                                 IF LEN(#mqttTopic) = #LEN_NULL THEN
                                   #statStatus := #ERR_MQTT_COMMAND_UNSUBSCRIBE_TOPIC_INVALID; // Set correct status that identifies error clearly
                                   #statSubfunctionStatus := #ERR_MQTT_COMMAND_UNSUBSCRIBE_TOPIC_INVALID; // Status or return value of called FBs, FCs and system blocks
                                   #statFBErrorState := #statFBState; // Set error state number for diagnostic 
                                   #statErrorUserCleared := TRUE;
                                 ELSE // All ok
                                   //Add two Byte for Paket ID:
                                   #statSendPaketTotalRemLen := #statSendPaketTotalRemLen + #TWO_BYTE_LEN_INFO;
                                   //add unsubscribe  topic len
                                   FOR #tempLoopCounter := #FIRST_CHARACTER TO LEN(#mqttTopic) DO
                                     "LMQTT_ConvertToUtf8"(character     := #mqttTopic[#tempLoopCounter],
                                                           convertedUtf8 => #tempConvertedUtf8,
                                                           bytesUsed     => #tempBytesUsedUtf8,
                                                           error         => #tempErrorConvertUtf8,
                                                           status        => #tempStatusConvertUtf8);
                                     #statUnsubscribeTopicLenUtf8Encoded := #statUnsubscribeTopicLenUtf8Encoded + #tempBytesUsedUtf8;
                                   END_FOR;
                                   //Add len of topic plus len info
                                   #statSendPaketTotalRemLen := #statSendPaketTotalRemLen + #statUnsubscribeTopicLenUtf8Encoded + #TWO_BYTE_LEN_INFO;

                                   //Build Subscribe Telegram
                                   //Fixed Header - Write Paket Type
                                   #statSendBuffer[#statSendBufferPos] := #MQTT_MSG_TYPE_UNSUBSCRIBE;
                                   #statSendBufferPos += 1; // increment

                                   //Write Remaining Paket Len info 
                                   WHILE (#statSendPaketTotalRemLen > #DEFAULT_VALUE_ZERO)
                                   DO//See MQTT Spec for explanation of this calculation
                                     #statEncodedRemPaketLenAsByte := UDINT_TO_BYTE(#statSendPaketTotalRemLen MOD #SEND_LEN_MULTIPLIER_UDINT_128);
                                     #statSendPaketTotalRemLen := #statSendPaketTotalRemLen / #SEND_LEN_MULTIPLIER_UDINT_128;
                                     // if there are more data to encode, set the top bit of this byte
                                     IF #statSendPaketTotalRemLen > #DEFAULT_VALUE_ZERO
                                     THEN
                                       // Do this and continue while loop
                                       #statEncodedRemPaketLenAsByte := #statEncodedRemPaketLenAsByte OR UDINT_TO_BYTE(#SEND_LEN_MULTIPLIER_UDINT_128);
                                       #statSendBuffer[#statSendBufferPos] := #statEncodedRemPaketLenAsByte;
                                       #statSendBufferPos += 1;
                                     ELSE
                                       //do this and leave while loop
                                       #statSendBuffer[#statSendBufferPos] := #statEncodedRemPaketLenAsByte;
                                       #statSendBufferPos += 1;
                                     END_IF;
                                   END_WHILE;

                                   // Set Paket Id
                                   #tempWordForSliceAddress := UINT_TO_WORD(#statPaketId);
                                   #statSendBuffer[#statSendBufferPos] := #tempWordForSliceAddress.%B1; //MSB
                                   #statSendBufferPos += 1;
                                   #statSendBuffer[#statSendBufferPos] := #tempWordForSliceAddress.%B0; //LSB
                                   #statSendBufferPos += 1;

                                   //When all done, set encode to true
                                   #statPaketHeaderEncodeDone := TRUE;
                                 END_IF;
                               END_IF;

                               //Header Encoded - 
                               IF #statPaketHeaderEncodeDone = TRUE THEN
                                 //Unsubscribe Topic
                                 IF #statSendBufferPos <= #MAX_BUFFER_LEN_SEND - #TWO_BYTE_LEN_INFO THEN
                                   CASE #statUnsubscribeTopicEncodeState OF
                                     #FIRST_ENCODING:  // Statement section case 1
                                       //ADD len info into paket

                                       #tempWordForSliceAddress := UINT_TO_WORD(#statUnsubscribeTopicLenUtf8Encoded);
                                       #statSendBuffer[#statSendBufferPos] := #tempWordForSliceAddress.%B1; //MSB
                                       #statSendBufferPos += 1;
                                       #statSendBuffer[#statSendBufferPos] := #tempWordForSliceAddress.%B0; // LSB
                                       #statSendBufferPos += 1;

                                       FOR #tempLoopCounter := #statUnsubscribeTopicPos TO LEN(#mqttTopic) DO
                                         "LMQTT_ConvertToUtf8"(character     := #mqttTopic[#tempLoopCounter],
                                                               convertedUtf8 => #tempConvertedUtf8,
                                                               bytesUsed     => #tempBytesUsedUtf8,
                                                               error         => #tempErrorConvertUtf8,
                                                               status        => #tempStatusConvertUtf8);

                                         IF #statSendBufferPos + #tempBytesUsedUtf8 <= #MAX_BUFFER_LEN_SEND THEN
                                           #statUnsubscribeTopicPos += 1;
                                           CASE #tempBytesUsedUtf8 OF
                                             #UTF_1_BYTE_USED:  // Statement section case 1
                                               #statSendBuffer[#statSendBufferPos] := #tempConvertedUtf8.%B0;
                                               #statSendBufferPos += 1;
                                             #UTF_2_BYTE_USED:
                                               #statSendBuffer[#statSendBufferPos] := #tempConvertedUtf8.%B0;
                                               #statSendBufferPos += 1;
                                               #statSendBuffer[#statSendBufferPos] := #tempConvertedUtf8.%B1;
                                               #statSendBufferPos += 1;
                                             #UTF_3_BYTE_USED:  // Statement section case 2 to 4
                                               #statSendBuffer[#statSendBufferPos] := #tempConvertedUtf8.%B0;
                                               #statSendBufferPos += 1;
                                               #statSendBuffer[#statSendBufferPos] := #tempConvertedUtf8.%B1;
                                               #statSendBufferPos += 1;
                                               #statSendBuffer[#statSendBufferPos] := #tempConvertedUtf8.%B2;
                                               #statSendBufferPos += 1;
                                             ELSE  // Statement section ELSE
                                               ;
                                           END_CASE;
                                         ELSE
                                           //When buffer full
                                           #statUnsubscribeTopicEncodeState := #SUBSEQUENT_ENCODING;
                                           EXIT;
                                         END_IF;
                                       END_FOR;
                                       IF #statUnsubscribeTopicPos >= LEN(#mqttTopic) THEN
                                         #statUnsubscribeTopicEncodeState := #ENCODE_DONE;
                                       END_IF;

                                     #SUBSEQUENT_ENCODING:  // Statement section case 2 to 4
                                       FOR #tempLoopCounter := #statUnsubscribeTopicPos TO LEN(#mqttTopic) DO

                                         "LMQTT_ConvertToUtf8"(character     := #mqttTopic[#tempLoopCounter],
                                                               convertedUtf8 => #tempConvertedUtf8,
                                                               bytesUsed     => #tempBytesUsedUtf8,
                                                               error         => #tempErrorConvertUtf8,
                                                               status        => #tempStatusConvertUtf8);
                                         IF #statSendBufferPos + #tempBytesUsedUtf8 <= #MAX_BUFFER_LEN_SEND THEN
                                           #statUnsubscribeTopicPos += 1;
                                           CASE #tempBytesUsedUtf8 OF
                                             #UTF_1_BYTE_USED:  // Statement section case 1
                                               #statSendBuffer[#statSendBufferPos] := #tempConvertedUtf8.%B0;
                                               #statSendBufferPos += 1;
                                             #UTF_2_BYTE_USED:
                                               #statSendBuffer[#statSendBufferPos] := #tempConvertedUtf8.%B0;
                                               #statSendBufferPos += 1;
                                               #statSendBuffer[#statSendBufferPos] := #tempConvertedUtf8.%B1;
                                               #statSendBufferPos += 1;
                                             #UTF_3_BYTE_USED:  // Statement section case 2 to 4
                                               #statSendBuffer[#statSendBufferPos] := #tempConvertedUtf8.%B0;
                                               #statSendBufferPos += 1;
                                               #statSendBuffer[#statSendBufferPos] := #tempConvertedUtf8.%B1;
                                               #statSendBufferPos += 1;
                                               #statSendBuffer[#statSendBufferPos] := #tempConvertedUtf8.%B2;
                                               #statSendBufferPos += 1;
                                             ELSE  // Statement section ELSE
                                               ;
                                           END_CASE;
                                         ELSE
                                           //When buffer full
                                           EXIT;
                                         END_IF;
                                       END_FOR;
                                       IF #statUnsubscribeTopicPos >= LEN(#mqttTopic) THEN
                                         #statUnsubscribeTopicEncodeState := #ENCODE_DONE;
                                       END_IF;
                                     ELSE  // Skip when Done
                                       ;
                                   END_CASE;
                                 END_IF;

                                 //set Sendlen for TSendC Block
                                 #statTsendcLen := #statSendBufferPos; // Buffer pos equals amount of elements in send array
                                 //reset buffer pos
                                 #statSendBufferPos := 0;
                                 //enable Send Req
                                 #statTsendcReq := TRUE;
                                 //Set Watchdog
                                 #statEnableTimerCommandWatchdog := TRUE;
                                 //wait for send to be done
                                 #statMqttCommandState := #MQTT_COMMAND_STATE_SEND_UNSUBSCRIBE;
                               END_IF;
                             END_IF;
                           END_REGION UNSUBSCRIBE_FROM_TOPIC

                         #MQTT_COMMAND_STATE_SEND_UNSUBSCRIBE:
                           REGION SEND_UNSUBSCRIBE_WAIT_FOR_RESPONSE
                             //check tsend status
                             IF NOT #tempTsendcBusy AND #tempTsendcStatus = #TSENDC_JOB_DONE THEN
                               IF (#statUnsubscribeTopicEncodeState = #ENCODE_DONE) THEN
                                 //Encoding done all sent
                                 #statPaketHeaderEncodeDone := FALSE;
                               ELSE
                                 // More to Encode and send
                                 #statEnableTimerCommandWatchdog := FALSE;
                                 #statMqttCommandState := #MQTT_COMMAND_STATE_BUILD_UNSUBSCRIBE;
                               END_IF;
                             END_IF;
                             // Wait for timeout
                             IF #instTimerCommandWatchdog.Q THEN
                               #statEnableTimerCommandWatchdog := FALSE;
                               #statStatus := #ERR_MQTT_COMMAND_SEND_TIMEOUT; // Set correct status that identifies error clearly
                               #statSubfunctionStatus := #ERR_MQTT_COMMAND_SEND_TIMEOUT; // Status or return value of called FBs, FCs and system blocks
                               #statFBErrorState := #statFBState; // Set error state number for diagnostic 
                               #statErrorAutoCleared := TRUE;
                               #statMqttCommandState := #MQTT_COMMAND_STATE_NO_PROCESSING;
                             END_IF;
                             //Check Unsubscribe ACK paket
                             CASE #tempMqttUnSubAckRcv OF
                               #NO_RESPONSE:  // Statement section case 1
                                 ;
                               #RESPONSE_GOOD:  // Statement section case 2 to 4
                                 //disable watchdog
                                 #statEnableTimerCommandWatchdog := FALSE;
                                 //Encoding done all sent
                                 #statPaketHeaderEncodeDone := FALSE;
                                 // Job done
                                 #statDone := TRUE;
                                 #statMqttCommandState := #MQTT_COMMAND_STATE_NO_PROCESSING;
                                 // Set Status back to connected
                                 #statStatus := #STATUS_JOB_EXECUTED;
                               #RESPONSE_PAKET_ID_INVALID:
                                 #statStatus := #ERR_MQTT_PAKET_ID_INVALID; // Set correct status that identifies error clearly
                                 #statSubfunctionStatus := #ERR_MQTT_PAKET_ID_INVALID; // Status or return value of called FBs, FCs and system blocks
                                 #statFBErrorState := #statFBState; // Set error state number for diagnostic 
                                 #statErrorAutoCleared := TRUE;
                                 #statMqttCommandState := #MQTT_COMMAND_STATE_NO_PROCESSING;
                             END_CASE;
                           END_REGION SEND_UNSUBSCRIBE_WAIT_FOR_RESPONSE

                         #MQTT_COMMAND_STATE_SEND_PING:
                           REGION SEND_PING
                             //Set Status
                             #statStatus := #STATUS_MQTT_PING;
                             IF #tempTsendcBusy = FALSE // when tsendC is ready
                               AND #tempTsendcDone = FALSE // tsendC did not finish in this cycle
                               AND #statTsendcReq = FALSE // TsendC request was not already requested by pub ack msg
                             THEN
                               //Init
                               #statSendBufferPos := 0;
                               #statSendBuffer[#statSendBufferPos] := #MQTT_MSG_TYPE_PING;
                               #statSendBufferPos += 1;
                               //Remaining Lenght (must be 0)
                               #statSendBuffer[#statSendBufferPos] := 0;
                               #statSendBufferPos += 1;
                               #statTsendcLen := #statSendBufferPos;
                               //Start send request
                               #statTsendcReq := TRUE;
                               //Start watchdoc
                               #statEnableTimerCommandWatchdog := true;
                               //Next state
                               #statMqttCommandState := #MQTT_COMMAND_STATE_PING_RESP;
                             END_IF;
                           END_REGION MQTT_COMMAND_SEND_PING

                         #MQTT_COMMAND_STATE_PING_RESP:
                           REGION WAIT_FOR_PING_RESP
                             //Check, if Edge of Publish comes while ping
                             IF #tempCommandInput > 0 AND NOT #statCommandInputOld THEN
                               #statCommandInputBackup := #tempCommandInput;
                               #statCommandInputOld := true;
                             END_IF;
                             //check watchdog status
                             IF #instTimerCommandWatchdog.Q THEN
                               #statEnableTimerCommandWatchdog := FALSE;
                               #statStatus := #ERR_MQTT_COMMAND_SEND_TIMEOUT; // Set correct status that identifies error clearly
                               #statSubfunctionStatus := #ERR_MQTT_COMMAND_SEND_TIMEOUT; // Status or return value of called FBs, FCs and system blocks
                               #statFBErrorState := #statFBState; // Set error state number for diagnostic 
                               #statErrorAutoCleared := TRUE;
                               #statMqttCommandState := #MQTT_COMMAND_STATE_NO_PROCESSING;
                             END_IF;
                             //Check PingRsp paket
                             CASE #tempMqttPingRspRcv OF
                               #NO_RESPONSE:  // Statement section case 1
                                 ;
                               #RESPONSE_GOOD:
                                 //disable watchdog
                                 #statEnableTimerCommandWatchdog := FALSE;
                                 //Go to no processing
                                 #statMqttCommandState := #MQTT_COMMAND_STATE_NO_PROCESSING;
                                 //set Status
                                 #statStatus := #STATUS_MQTT_CONNECTED;
                                 IF #statCommandInputBackup <> 0 THEN
                                   #statMqttCommandState := BYTE_TO_DINT(#statCommandInputBackup);
                                   #statCommandInputBackup := 0;
                                   #statCommandInputOld := false;
                                 END_IF;
                             END_CASE;
                           END_REGION MQTT_COMMAND_PING_RESP
                         ELSE  // Statement section ELSE
                           REGION ERROR_MULTIPLE_INPUT
                             #statMqttCommandState := #MQTT_COMMAND_STATE_NO_PROCESSING; // reset back to idle
                             #statStatus := #ERR_MQTT_COMMAND_MULTIPLE_INPUT; // Set correct status that identifies error clearly
                             #statSubfunctionStatus := #ERR_MQTT_COMMAND_MULTIPLE_INPUT; // Status or return value of called FBs, FCs and system blocks
                             #statFBErrorState := #statFBState; // Set error state number for diagnostic 
                             #statErrorAutoCleared := TRUE;
                           END_REGION ERROR_MULTIPLE_INPUT 
                       END_CASE;
                     END_REGION

                     REGION CHECK_PING_TIMER
                       //If no job is running check if keepalive experied
                       IF #statMqttCommandState = #MQTT_COMMAND_STATE_NO_PROCESSING
                         AND #instMqttKeepAliveTimer.Q THEN
                         //reset the timer
                         RESET_TIMER(#instMqttKeepAliveTimer);
                         //go to ping state
                         #statMqttCommandState := #MQTT_COMMAND_STATE_SEND_PING;
                       END_IF;
                     END_REGION CHECK_PING_TIMER

                     //Edge detection "publish / subscribe/unsubscribe" input
                     #statPublishOld := #tempPublish;
                     #statSubscribeOld := #tempSubscribe;
                     #statUnsubscribeOld := #tempUnsubscribe;
                   END_REGION CONNECTED

                 ELSE   // Undefined state in state machine reached
                   #statStatus := #ERR_UNDEFINED_STATE;
                   #statErrorUserCleared := TRUE;
               END_CASE;

             END_REGION MQTT_STATE_MACHINE
           END_IF;
         END_REGION FB_OPERATING_MONITOR_TCP

       #FB_STATE_TCP_RECONNECTING:
         REGION FB_STATE_TCP_RECONNECTING
           IF #tempTsendcStatus = #TSENDC_EST_OK THEN
             #statErrorAutoCleared := FALSE;
             // Update edge detection
             #statPublishOld := #tempPublish;
             #statSubscribeOld := #tempSubscribe;
             #statUnsubscribeOld := #tempUnsubscribe;
             //Monitor Connection
             #statFBState := #FB_STATE_OPERATING_MONITOR_TCP;
             // Begin MQTT Connection
             #statMqttConnectState := #MQTT_CONNECT_STATE_BUILD_PAKET;
           END_IF;
         END_REGION FB_STATE_TCP_RECONNECTING
       #FB_STATE_DISABLING: // Disabling active
         REGION DISABLING FB
           //  Disabling, e.g. closing connections, etc.
           // When disabling is complete the bit #statDisablingCompleted must be set
           // When MQTT is connected, send disconnect
           IF #statMqttConnectState = #MQTT_CONNECT_STATE_CONNECTED THEN
             IF #statTsendcReq = TRUE THEN
               //Interrupt any existing send jobs
               #statTsendcReq := FALSE;
             ELSE
               // INIT
               #statSendBufferPos := 0;
               //Build fixed Header
               //Message Type
               #statSendBuffer[#statSendBufferPos] := #MQTT_MSG_TYPE_DISCONNECT;
               #statSendBufferPos += 1;
               //Remaining Length (must be O)
               #statSendBuffer[#statSendBufferPos] := #REMAINIG_LEN_0;
               #statSendBufferPos += 1;
               //send request
               #statTsendcLen := #statSendBufferPos;
               #statTsendcReq := TRUE;
               #statMqttConnectState := #MQTT_CONNECT_STATE_DISCONNECTED;
             END_IF;
           ELSE
             //Disable TCP Connection
             #statTsendcReq := FALSE;
             #statTsendcEnable := FALSE;
             #statEnableTimerCommandWatchdog := TRUE;
           END_IF;
           // When TCP connection is closed
           IF #tempTsendcStatus = #TSENDC_DISCONNECTED THEN
             #statEnableTimerCommandWatchdog := FALSE;
             #statDisablingCompleted := TRUE;
           ELSIF #instTimerCommandWatchdog.Q THEN
             #statEnableTimerCommandWatchdog := FALSE;
             #statDisablingCompleted := TRUE;
           END_IF;
         END_REGION DISABLING FB
       ELSE // Undefined state in state machine reached
         #statStatus := #ERR_UNDEFINED_STATE;
         #statErrorUserCleared := TRUE;
     END_CASE;
   END_REGION STATE_MACHINE

   REGION OUTPUTS
     // Write outputs
     IF (#statDisablingCompleted = TRUE) THEN
       // Reset outputs if disabling completed
       #statValid := FALSE;
       #statBusy := FALSE;
       #statError := FALSE;
       #statDone := FALSE;
       #statErrorUserCleared := FALSE;
       #statErrorAutoCleared := FALSE;
       #statStatus := #STATUS_NO_CALL;
       // Reset application specific outputs
       #statRcvMsgStatus := #MSG_DECODE_STATUS_NO_NEW_MSG;
       #statRcvMsgDataLen := 0;

     ELSIF (#statErrorUserCleared = TRUE) AND (#statError = FALSE) THEN
       // Error can only be cleared by user; rising edge at enable input is needed to continue 
       #statValid := FALSE;
       #statBusy := FALSE;
       #statDone := FALSE;
       #statError := TRUE;
       // Write diagnostics
       #diagnostics.status := #statStatus;
       #diagnostics.subfunctionStatus := #statSubfunctionStatus;
       #diagnostics.stateNumber := #statFBErrorState;
       // execution aborted --> set state no processing
       #statTsendcEnable := FALSE; // Terminate Connection, no reason keep it up.
       #statFBState := #FB_STATE_NO_PROCESSING;
       #statMqttConnectState := #MQTT_CONNECT_STATE_NO_PROCESSING;
       #statMqttCommandState := #MQTT_COMMAND_STATE_NO_PROCESSING;
       #statRcvMsgDecodeState := #MSG_DECODE_STATE_NO_PROCESSING;

     ELSIF (#statErrorAutoCleared = TRUE) AND (#statError = FALSE) THEN
       // Error can be reset by FB automatically
       #statValid := FALSE;
       #statBusy := TRUE;
       #statError := TRUE;
       #statDone := FALSE;

       // Write diagnostics
       #diagnostics.status := #statStatus;
       #diagnostics.subfunctionStatus := #statSubfunctionStatus;
       #diagnostics.stateNumber := #statFBErrorState;
       // Handling of autocleared error
       CASE #statStatus OF
           //Just signal error and reset autocleared error afterwards.
         #ERR_MQTT_PAKET_ID_INVALID, #ERR_MQTT_SUBACK_FAILURE, #ERR_MQTT_CONNECT_TIMEOUT,
         #ERR_MQTT_COMMAND_SEND_TIMEOUT, #ERR_MQTT_COMMAND_MULTIPLE_INPUT, #ERR_CNT_EXCEEDS_ARRAY_DIMENSION,
         #ERR_MQTT_COMMAND_PUBLISH_TOPIC_INVALID, #ERR_QOS_INVALID, #ERR_MQTT_COMMAND_SUBSCRIBE_TOPIC_INVALID:
           #statErrorAutoCleared := FALSE;

         ELSE  // Statement section ELSE
           ;
       END_CASE;

     ELSIF (#statErrorAutoCleared = FALSE) AND (#statErrorUserCleared = FALSE) AND (#statError = TRUE) THEN
       // If autocleared error is acknowledged
       #statValid := TRUE;
       #statBusy := TRUE;
       #statError := FALSE;
       #statDone := FALSE;

       //   this line  more detailed status information is used instead of "#STATUS_SUBSEQUENT_CALL"
       CASE #statStatus OF
         #ERR_TCP_RECONNECTING, #ERR_MQTT_CONNECT_TIMEOUT:  // Reconnecting ok, start Mqtt reconnnect
           //set status
           #statStatus := #STATUS_MQTT_CONNECTING;
           //in the following status codes status stays connected. 
         #ERR_MQTT_PAKET_ID_INVALID, #ERR_MQTT_SUBACK_FAILURE, #ERR_MQTT_COMMAND_SEND_TIMEOUT,
         #ERR_MQTT_COMMAND_MULTIPLE_INPUT, #ERR_CNT_EXCEEDS_ARRAY_DIMENSION, #ERR_MQTT_COMMAND_PUBLISH_TOPIC_INVALID,
         #ERR_QOS_INVALID, #ERR_MQTT_COMMAND_SUBSCRIBE_TOPIC_INVALID:
           #statStatus := #STATUS_MQTT_CONNECTED;
         ELSE  // Statement section ELSE
           ;
       END_CASE;
     END_IF;

     // Write static values to outputs
     #valid := #statValid;
     #busy := #statBusy;
     #error := #statError;
     #status := #statStatus;
     //block sets ENO automatically:
     //ENO := TRUE;
     //Write application specific static values to outputs
     #done := #statDone;
     #receivedMsgStatus := #statRcvMsgStatus;
     #receivedMsgDataLen := #statRcvMsgDataLen;
   END_REGION OUTPUTS
END_FUNCTION_BLOCK

FUNCTION "INPUTS" : Void   // FC25, SCL
{ S7_Optimized_Access := 'TRUE' }
VERSION : 0.1
// stored: AutoNumber true, IsIECCheckEnabled false, SetENOAutomatically false, UDAEnableTagReadback false
   VAR_TEMP
      Barcode_Inbound : Array[1..16] of Char;
      Barcode_Outbound : Array[1..16] of Char;
      Empty_code : Array[1..16] of Char;
   END_VAR
BEGIN
   REGION INBOUND CONVEYOR
       "Control_DB".Inbound_Cnv.Inputs."Pallet Detect 1" := NOT "Inbound Conveyor - Back Sensor";
       "Control_DB".Inbound_Cnv.Inputs."Pallet Detect 2" := NOT "Inbound Conveyor - Front Sensor";
       "Control_DB".Inbound_Cnv.Inputs."Fork Lift Detect":= "Fork Lift Detect_Inbound";
   END_REGION

   REGION OUTBOUND CONVEYOR
       "Control_DB".Outbound_Cnv.Inputs."Pallet Detect" := "Outbound Conveyor";
       "Control_DB".Outbound_Cnv.Inputs."Fork Lift Detect" := "Fork Lift Detect_Outbound";
   END_REGION

   REGION EXTRACTOR CONVEYOR
       "Control_DB".ECnv_Control.Inputs."Pallet Detect 1" := "Pallet in Position Front VTD";
       "Control_DB".ECnv_Control.Inputs."Pallet Detect 2" := "Pallet in Position Rear VTD";
       "Control_DB".ECnv_Control.Inputs.Sdetect1 := "Shuttle in Position Front VTD";
       "Control_DB".ECnv_Control.Inputs.Sdetect2 := "Shuttle in Position Rear VTD";
   END_REGION

   REGION BUFFER CONVEYOR
       //BUFFER CONVEYOR LEVEL 1
       "Control_DB".LCnv_Control[1].Inputs."Pallet Detect 1" := "Buffer Conveyor 1 - Pallet present 1";
       "Control_DB".LCnv_Control[1].Inputs."Pallet Detect 2" := "Buffer Conveyor 1 - Pallet present 2";
       "Control_DB".LCnv_Control[1].Inputs."Pallet Detect 3" := "Buffer Conveyor 1 - Pallet present 3";
       "Control_DB".LCnv_Control[1].Inputs.Sdetect1 := "Buffer Conveyor 1 - Shuttle present 1";
       "Control_DB".LCnv_Control[1].Inputs.Sdetect2 := "Buffer Conveyor 1 - Shuttle present 2";
       "Control_DB".LCnv_Control[1].Inputs.SftyPinUp := "Buffer Conveyor 1 - Safety Pin Up";
       "Control_DB".LCnv_Control[1].Inputs.SftyPinDown := "Buffer Conveyor 1 - Safety Pin Down";
       //BUFFER CONVEYOR LEVEL 2
       "Control_DB".LCnv_Control[2].Inputs."Pallet Detect 1" := "Buffer Conveyor 2 - Pallet present 1";
       "Control_DB".LCnv_Control[2].Inputs."Pallet Detect 2" := "Buffer Conveyor 2 - Pallet present 2";
       "Control_DB".LCnv_Control[2].Inputs."Pallet Detect 3" := "Buffer Conveyor 2 - Pallet present 3";
       "Control_DB".LCnv_Control[2].Inputs.Sdetect1 := "Buffer Conveyor 2 - Shuttle present 1";
       "Control_DB".LCnv_Control[2].Inputs.Sdetect2 := "Buffer Conveyor 2 - Shuttle present 2";
       "Control_DB".LCnv_Control[2].Inputs.SftyPinUp := "Buffer Conveyor 2 - Safety Pin Up";
       "Control_DB".LCnv_Control[2].Inputs.SftyPinDown := "Buffer Conveyor 2 - Safety Pin Down";
       //BUFFER CONVEYOR LEVEL 3
       "Control_DB".LCnv_Control[3].Inputs."Pallet Detect 1" := "Buffer Conveyor 3 - Pallet present 1";
       "Control_DB".LCnv_Control[3].Inputs."Pallet Detect 2" := "Buffer Conveyor 3 - Pallet present 2";
       "Control_DB".LCnv_Control[3].Inputs."Pallet Detect 3" := "Buffer Conveyor 3 - Pallet present 3";
       "Control_DB".LCnv_Control[3].Inputs.Sdetect1 := "Buffer Conveyor 3 - Shuttle present 1";
       "Control_DB".LCnv_Control[3].Inputs.Sdetect2 := "Buffer Conveyor 3 - Shuttle present 2";
       "Control_DB".LCnv_Control[3].Inputs.SftyPinUp := "Buffer Conveyor 3 - Safety Pin Up";
       "Control_DB".LCnv_Control[3].Inputs.SftyPinDown := "Buffer Conveyor 3 - Safety Pin Down";
   END_REGION

   REGION VTD
       "Control_DB".VTD_Control.Inputs.Upper_limit := "Upper Ultimate";
       "Control_DB".VTD_Control.Inputs.Lower_Limit := "Lower Ultimate";
       "Control_DB".VTD_Control.Inputs.Level_Detect1 := "Docking Sensor Front";
       "Control_DB".VTD_Control.Inputs.Level_Detect2 := "Docking Sensor Rear";
       "Control_DB".VTD_Control.Inputs.Ultimate_Slow := "Slowdown";
       "Control_DB".VTD_Control.Inputs.Ultimate_Creep := "Creep speed";
       "Control_DB".VTD_Control.Inputs.LPL_Extended := "Locking Pins Extended left";
       "Control_DB".VTD_Control.Inputs.LPR_Extended := "Locking Pins Extended Right";
       "Control_DB".VTD_Control.Inputs.LPL_Retracted := "Locking Pins Retracted left";
       "Control_DB".VTD_Control.Inputs.LPR_Retracted := "Locking Pins Retracted Right";
   END_REGION

   REGION POPUP CONVEYORS
       "Control_DB".PopUp_Cnv[1].Inputs."Lift Up" := "PopUp Conveyor 1 - Sensor Up";
       "Control_DB".PopUp_Cnv[1].Inputs."Lift Down" := "PopUp Conveyor 1 - Sensor Down";
       "Control_DB".PopUp_Cnv[2].Inputs."Lift Up" := "PopUp Conveyor 2 - Sensor Up";
       "Control_DB".PopUp_Cnv[2].Inputs."Lift Down" := "PopUp Conveyor 2 - Sensor Down";
       "Control_DB".PopUp_Cnv[3].Inputs."Lift Up" := "PopUp Conveyor 3 - Sensor Up";
       "Control_DB".PopUp_Cnv[3].Inputs."Lift Down" := "PopUp Conveyor 3 - Sensor Down";
       "Control_DB".PopUp_Cnv[4].Inputs."Lift Up" := "PopUp Conveyor 4 - Sensor Up";
       "Control_DB".PopUp_Cnv[4].Inputs."Lift Down" := "PopUp Conveyor 4 - Sensor Down";
   END_REGION

   REGION VFD HARDWARE ID
       //Buffer conveyors
       "Settings_DB".LCnv_Settings[1].G120_Hardware_ID := "Buffer_Level1~PROFINET_interface~Standard_telegram_1";
       "Settings_DB".LCnv_Settings[2].G120_Hardware_ID := "Buffer_Level2~PROFINET_interface~Standard_telegram_1";
       "Settings_DB".LCnv_Settings[3].G120_Hardware_ID := "Buffer_Level3~PROFINET_interface~Standard_telegram_1";
       //Extractor conveyor
       "Settings_DB".ECnv_Settings.G120_Hardware_ID := "VTD_Coveyor~PROFINET_interface~Standard_telegram_1";
       //IO Conveyors
       "Settings_DB".Inbound_Cnv_Settings.G120_Hardware_ID := "Roller_Inbound~PROFINET_interface~Standard_telegram_1";
       "Settings_DB".Outbound_Cnv_Settings.G120_Hardware_ID := "Roller_Outbound~PROFINET_interface~Standard_telegram_1";
       //PopUp conveyor 1
       "Settings_DB".PopUp_Cnv_Settings[1].Roller_G120_Hardware_ID := "Roller_PopUp1~PROFINET_interface~Standard_telegram_1";
       "Settings_DB".Pick_Cnv_Settings.G120_Hardware_ID := "Chain1~PROFINET_interface~Standard_telegram_1";
       "Settings_DB".PopUp_Cnv_Settings[1].Lift_G120_Hardware_ID := "Lift_PopUp1~PROFINET_interface~Standard_telegram_1";
       //PopUp conveyor 2
       "Settings_DB".PopUp_Cnv_Settings[2].Roller_G120_Hardware_ID := "Roller_PopUp2~PROFINET_interface~Standard_telegram_1";
       "Settings_DB".PopUp_Cnv_Settings[2].Chain_G120_Hardware_ID := "Chain2~PROFINET_interface~Standard_telegram_1";
       "Settings_DB".PopUp_Cnv_Settings[2].Lift_G120_Hardware_ID := "Lift_PopUp2~PROFINET_interface~Standard_telegram_1";
       //PopUp conveyor 3
       "Settings_DB".PopUp_Cnv_Settings[3].Roller_G120_Hardware_ID := "Roller_PopUp3~PROFINET_interface~Standard_telegram_1";
       "Settings_DB".PopUp_Cnv_Settings[3].Chain_G120_Hardware_ID := "Chain3~PROFINET_interface~Standard_telegram_1";
       "Settings_DB".PopUp_Cnv_Settings[3].Lift_G120_Hardware_ID := "Lift_PopUp3~PROFINET_interface~Standard_telegram_1";
       //PopUp conveyor 4
       "Settings_DB".PopUp_Cnv_Settings[4].Roller_G120_Hardware_ID := "Roller_PopUp4~PROFINET_interface~Standard_telegram_1";
       "Settings_DB".PopUp_Cnv_Settings[4].Lift_G120_Hardware_ID := "Lift_PopUp4~PROFINET_interface~Standard_telegram_1";
   END_REGION

   REGION LEUZE/SICK BARCODE LECTORS
       #Barcode_Inbound[1] := "In Lector_Data - Byte 1";
       #Barcode_Inbound[2] := "In Lector_Data - Byte 2";
       #Barcode_Inbound[3] := "In Lector_Data - Byte 3";
       #Barcode_Inbound[4] := "In Lector_Data - Byte 4";
       #Barcode_Inbound[5] := "In Lector_Data - Byte 5";
       #Barcode_Inbound[6] := "In Lector_Data - Byte 6";
       #Barcode_Inbound[7] := "In Lector_Data - Byte 7";
       #Barcode_Inbound[8] := "In Lector_Data - Byte 8";
       #Barcode_Inbound[9] := "In Lector_Data - Byte 9";
       #Barcode_Inbound[10] := "In Lector_Data - Byte 10";
       #Barcode_Inbound[11] := "In Lector_Data - Byte 11";
       #Barcode_Inbound[12] := "In Lector_Data - Byte 12";
       #Barcode_Inbound[13] := "In Lector_Data - Byte 13";
       #Barcode_Inbound[14] := "In Lector_Data - Byte 14";
       #Barcode_Inbound[15] := "In Lector_Data - Byte 15";
       #Barcode_Inbound[16] := "In Lector_Data - Byte 16";

       #Barcode_Outbound[1] := "Out Lector_Data - Byte 1";
       #Barcode_Outbound[2] := "Out Lector_Data - Byte 2";
       #Barcode_Outbound[3] := "Out Lector_Data - Byte 3";
       #Barcode_Outbound[4] := "Out Lector_Data - Byte 4";
       #Barcode_Outbound[5] := "Out Lector_Data - Byte 5";
       #Barcode_Outbound[6] := "Out Lector_Data - Byte 6";
       #Barcode_Outbound[7] := "Out Lector_Data - Byte 7";
       #Barcode_Outbound[8] := "Out Lector_Data - Byte 8";
       #Barcode_Outbound[9] := "Out Lector_Data - Byte 9";
       #Barcode_Outbound[10] := "Out Lector_Data - Byte 10";
       #Barcode_Outbound[11] := "Out Lector_Data - Byte 11";
       #Barcode_Outbound[12] := "Out Lector_Data - Byte 12";
       #Barcode_Outbound[13] := "Out Lector_Data - Byte 13";
       #Barcode_Outbound[14] := "Out Lector_Data - Byte 14";
       #Barcode_Outbound[15] := "Out Lector_Data - Byte 15";
       #Barcode_Outbound[16] := "Out Lector_Data - Byte 16";




       IF "Control_DB".OutBarcode_Station.Running AND #Barcode_Outbound <> "Control_DB".OutBarcode_Station.Barcode_Old THEN
           "Control_DB".Outbound_Cnv.Inputs.Barcode := "CharsArrayToString"(CharsArray := #Barcode_Outbound, Lenght := 16);
           "Control_DB".OutBarcode_Station.Barcode_Old := #Barcode_Outbound;
       ELSE
           "Control_DB".OutBarcode_Station.Barcode := '';
       END_IF;

       IF "Control_DB".VTDBarcode_Station.Running AND "SICK_Barcode_DB".Result <> "Control_DB".VTDBarcode_Station.Barcode_Old THEN
           "Control_DB".VTD_Control.Inputs."Barcode 1" := "SICK_Barcode_DB".Result;
           // "Control_DB".VTD_Control.Inputs."Barcode 2'" := SICK_Barcode_DB".Result;
           "Control_DB".VTDBarcode_Station.Barcode_Old := "SICK_Barcode_DB".Result;
       ELSE
           "Control_DB".VTD_Control.Inputs."Barcode 1" :=
           "Control_DB".VTD_Control.Inputs."Barcode 2'" :='';
       END_IF;

       // IF "Reset_All" THEN
       //     "Control_DB".InBarcode_Station."Reading Gate number OLD" := '';
       //     "Control_DB".OutBarcode_Station.Barcode_Old := #Empty_code;
       //     "Control_DB".VTD_Control.Inputs."Barcode 1" := 
       //     "Control_DB".VTD_Control.Inputs."Barcode 2'" := '';
       // END_IF;
   END_REGION

   REGION WEIGTH STATION
       "SB_Alarm"."LC overload in operation range" := "SB Status Group 1".%X0;
       "SB_Alarm"."LC Mix" := "SB Status Group 1".%X1;
       "SB_Alarm"."Application defined 1" := "SB Status Group 1".%X2;
       "SB_Alarm"."Application defined 2" := "SB Status Group 1".%X3;
       "SB_Alarm"."Application defined 3" := "SB Status Group 1".%X4;
       "SB_Alarm"."Application defined 4" := "SB Status Group 1".%X5;
       "SB_Alarm"."Application defined 5" := "SB Status Group 1".%X6;
       "SB_Alarm"."Application defined 7" := "SB Status Group 1".%X7;
       "SB_Alarm"."Rate of change error" := "SB Status Group 1".%X8;
       "SB_Alarm"."Communication error" := "SB Status Group 1".%X9;
       "SB_Alarm"."Over / under voltage" := "SB Status Group 1".%X10;
       "SB_Alarm"."Weight drift" := "SB Status Group 1".%X11;
       "SB_Alarm".Breach := "SB Status Group 1".%X12;
       "SB_Alarm"."Calibration expired" := "SB Status Group 1".%X13;
       "SB_Alarm"."Over Current" := "SB Status Group 1".%X14;
       "SB_Alarm"."LC overload in normal range" := "SB Status Group 1".%X15;

       "SB_RedAlarm"."Zero out of range" := "SB Status Group 2".%X0;
       "SB_RedAlarm"."Symetry errors" := "SB Status Group 2".%X1;
       "SB_RedAlarm"."LC Temperature out of normal temperature" := "SB Status Group 2".%X2;
       "SB_RedAlarm"."Weights and measures failure" := "SB Status Group 2".%X3;
       "SB_RedAlarm"."Foreign device detected" := "SB Status Group 2".%X4;
       "SB_RedAlarm"."Test mode" := "SB Status Group 2".%X5;
       "SB_RedAlarm"."LC temperature out of operatio" := "SB Status Group 2".%X6;
       "SB_RedAlarm"."LC parameters block checksum error" := "SB Status Group 2".%X7;
       "SB_RedAlarm"."Calibration error" := "SB Status Group 2".%X8;
       "SB_RedAlarm"."Out of A/D range over/under" := "SB Status Group 2".%X9;
       "SB_RedAlarm"."Checksu failure" := "SB Status Group 2".%X10;
       "SB_RedAlarm"."Weight blocked" := "SB Status Group 2".%X11;
       "SB_RedAlarm"."LC Missing" := "SB Status Group 2".%X12;
       "SB_RedAlarm"."Customer-defined overload" := "SB Status Group 2".%X13;
       "SB_RedAlarm"."Customer-defined underload" := "SB Status Group 2".%X14;
   END_REGION

   REGION PICK STATION
       "Control_DB".Pick_Station.Cnv_Occupied := NOT "Pick Station";
       "Control_DB".Pick_Station.PushButton := "PushButton Pick Station";
       "Control_DB".Pick_Station.LightGuard := NOT "LighGuard_Cut-Off Path 01";
   END_REGION
END_FUNCTION

FUNCTION_BLOCK "VTD_HMI_FB"   // FB14, SCL
{ S7_Optimized_Access := 'TRUE' }
VERSION : 0.1
// stored: AutoNumber true, IsIECCheckEnabled false, IsRetainMemResEnabled false, MemoryReserve 100, SetENOAutomatically false, UDAEnableTagReadback false
BEGIN
   //CHARGE DATA
   "R_TRIG_DB_6"(CLK:="Screen_DB".Charge_VTD_Commands);

   IF "R_TRIG_DB_6".Q THEN
       "VTD_Mode_Change_HMI_Tag" := "Control_DB".VTD_Control.Mode;
       "VTD_Enable_HMI_Tag" := "Control_DB".VTD_Control.Instruction.Enable;
       "IEC_Timer_0_DB_2_IN" := TRUE;
   END_IF;
   "IEC_Timer_0_DB_2".TON(IN := "IEC_Timer_0_DB_2_IN",
                          PT := T#1S);
   IF "IEC_Timer_0_DB_2".Q THEN
       "IEC_Timer_0_DB_2_IN" := FALSE;
       "Screen_DB".Charge_VTD_Commands := 0;
   END_IF;

   REGION VTD HMI Assignments
       // Statement section REGION

       //Status
       "VTD_Error_Feedback_HMI_Tag" := "Control_DB".VTD_Control.Error;
       "VTD_Warning_Feedback_HMI_Tag" := "Control_DB".VTD_Control.Warning <> 0;
       "VTD_Enabled_Feedback_HMI_Tag" := "Control_DB".VTD_Control.Enabled;
       "VTD_Stopped_Feedback_HMI_Tag" := "Control_DB".VTD_Control.Stopped;
       "VTD_Running_Feedback_HMI_Tag" := "Control_DB".VTD_Control.Running;
       "VTD_Docked_Feedback_HMI_Tag" := "Control_DB".VTD_Control.Docked;
       "VTD_Current_Task_Type_Feedback_HMI_Tag" := "Control_DB".VTD_Control.Current_Task_Type;
       "VTD_Current_Task_ID_Feedback_HMI_Tag" := "Control_DB".VTD_Control.Current_Task_ID;
       "VTD_Current_Level_Feedback_HMI_Tag" := "Control_DB".VTD_Control.Current_Level;
       "VTD_LP_State_Feedback_HMI_Tag" := "Control_DB".VTD_Control.LP_State;
       "VTD_Pallet_Loaded_Feedback_HMI_Tag" := "Control_DB".VTD_Control.Pallet_Loaded;
       "VTD_Shuttle_Loaded_Feedback_HMI_Tag" := "Control_DB".VTD_Control.Shuttle_Loaded;
       "VTD_SM_State_Feedback_HMI_Tag" := "Control_DB".VTD_Control.SM_State;
       "VTD_LE_Error_Feedback_HMI_Tag" := "LE_Status".%X0;
       "VTD_AE_Error_Feedback_HMI_Tag" := "AE_Status_2".%X15;
       "VTD_Encoder_Delta_Feedback_HMI_Tag" := "Control_DB".VTD_Control.Encoder_Delta;
       "VTD_AE_Feedback_HMI_Tag" := "Control_DB".VTD_Control.AE;
       "VTD_LE_Feedback_HMI_Tag" := "Control_DB".VTD_Control.LE;

       "VTD_Progress_HMI_Tag" := "Control_DB".VTD_Control.LE;

       //Inputs
       "VTD_Upper_Limet_HMI_Tag" := "Upper Ultimate";
       "VTD_Lower_Limit_HMI_Tag" := "Lower Ultimate";
       "VTD_Lower_Overtravel_HMI_Tag" := "Overtravel Lower Limit - CH1";
       "VTD_Upper_Overtravel_HMI_Tag" := "Overtravel Upper Limit - CH1";
       "VTD_Level_Detect1_HMI_Tag" := "Docking Sensor Front";
       "VTD_Level_Detect2_HMI_Tag" := "Docking Sensor Rear";
       "VTD_Ultimate_Slow_HMI_Tag" := "Slowdown";
       "VTD_Ultimate_Creep_HMI_Tag" := "Creep speed";
       "VTD_LPL_Extended_HMI_Tag" := "Locking Pins Extended left";
       "VTD_LPR_Extended_HMI_Tag" := "Locking Pins Extended Right";
       "VTD_LPL_Retracted_HMI_Tag" := "Locking Pins Retracted left";
       "VTD_LPR_Retracted_HMI_Tag" := "Locking Pins Retracted Right";

       //Instruction
       IF "HMI_DB".ScreenNo = 1 AND NOT "Screen_DB".Charge_VTD_Commands THEN
           "Control_DB".VTD_Control.Instruction.Reset := "VTD_Reset_HMI_Tags";
           "Control_DB".VTD_Control.Instruction.Execulte := "VTD_Execute";
           "Control_DB".VTD_Control.Instruction.Mode_Change := "VTD_Mode_Change_HMI_Tag";
           "Control_DB".VTD_Control.Instruction.Enable := "VTD_Enable_HMI_Tag";

           IF "Control_DB".VTD_Control.Mode <> 3 THEN

               // "Control_DB".VTD_Control.Instruction.Stop := "VTD_Stop_HMI_Tag";
               "Control_DB".VTD_Control.Instruction.Pallet_Type := "VTD_Pallet_Type_HMI_Tag";
               "Control_DB".VTD_Control.Instruction.Task_ID := "VTD_Task_ID_HMI_Tag";
               "Control_DB".VTD_Control.Instruction.Move_To_Level := "VTD_Move_To_Level_HMI_Tag";
               "Control_DB".VTD_Control.Instruction.Manual_Up := "VTD_Manual_Up_HMI_Tag";
               "Control_DB".VTD_Control.Instruction.Manual_Down := "VTD_Manual_Down_HMI_Tag";
               "Control_DB".VTD_Control.Instruction.Manual_LP_Retract := "VTD_Manual_LP_Retract_HMI_Tags";
               "Control_DB".VTD_Control.Instruction.Manual_LP_Extend := "VTD_Manual_LP_Extend_HMI_Tags";
               "Control_DB".VTD_Control.Instruction.Start_Teach := "VTD_Start_Teach_HMI_Tags";
           END_IF;
       END_IF;
   END_REGION
END_FUNCTION_BLOCK

FUNCTION_BLOCK "Conveyor_HMI_FB"   // FB13, SCL
{ S7_Optimized_Access := 'TRUE' }
VERSION : 0.1
// stored: AutoNumber true, IsIECCheckEnabled false, IsRetainMemResEnabled false, MemoryReserve 100, SetENOAutomatically false, UDAEnableTagReadback false
   VAR_TEMP
      i : UInt;
      J : UInt;
   END_VAR
BEGIN
   REGION Assign Conveyor 1
       REGION Charge DATA
           IF "CNV_ID_HMI_Tag" = "CNV_ID_HMI_Tag(1)" THEN
               //CNV 1
               "Same_Cnv" := TRUE;

               "Enable_HMI_Tag" := 0;
               "Mode_Change_HMI_Tag" := 0;
               "Task_ID_HMI_Tag" := 0;
               "Transfer_To_ID_HMI_Tag" := 0;
               "Transfer_From_ID_HMI_Tag" := 0;
               //Sensors
               "HMI_CNV_Pallet Detect 1" := 0;
               "HMI_CNV_Pallet Detect 2" := 0;
               "HMI_CNV_Pallet Detect 3" := 0;
               "HMI_CNV_Sdetect1" := 0;
               "HMI_CNV_Sdetect2" := 0;
               "HMI_CNV_SftyPinUp" := 0;
               "HMI_CNV_SftyPinDown" := 0;

               //Feedback
               "Mode_HMI_Feedback_Tag" := 0;
               "Enabled_HMI_Feedback_Tag" := 0;
               "Error_HMI_Feedback_Tag" := 0;
               "Warning_HMI_Feedback_Tag" := 0;
               "Stopped_HMI_Feedback_Tag" := 0;
               "Running_HMI_Feedback_Tag" := 0;
               "Ready_For_Task_HMI_Feedback_Tag" := 0;
               "Cnv_Occupied_HMI_Feedback_Tag" := 0;
               "Shuttle_in_place_HMI_Feedback_Tag" := 0;
               "Current_Task_Type_HMI_Feedback_Tag" := 0;
               "Current_Task_ID_HMI_Feedback_Tag" := 0;
               "SM_State_HMI_Feedback_Tag" := 0;
               "Motor_Speed_Requested_HMI_Feedback_Tag" := 0;
               "Motor_Speed_Actual_HMI_Feedback_Tag" := 0;

               //CNV 2
               "Enable_HMI_Tag(1)" := 0;
               "Mode_Change_HMI_Tag(1)" := 0;
               "Task_ID_HMI_Tag(1)" := 0;
               "Transfer_To_ID_HMI_Tag(1)" := 0;
               "Transfer_From_ID_HMI_Tag(1)" := 0;
               //Sensors
               "HMI_CNV_Pallet Detect 1(1)" := 0;
               "HMI_CNV_Pallet Detect 2(1)" := 0;
               "HMI_CNV_Pallet Detect 3(1)" := 0;
               "HMI_CNV_Sdetect1(1)" := 0;
               "HMI_CNV_Sdetect2(1)" := 0;
               "HMI_CNV_SftyPinUp(1)" := 0;
               "HMI_CNV_SftyPinDown(1)" := 0;

               //Feedback
               "Mode_HMI_Feedback_Tag(1)" := 0;
               "Enabled_HMI_Feedback_Tag(1)" := 0;
               "Error_HMI_Feedback_Tag(1)" := 0;
               "Warning_HMI_Feedback_Tag(1)" := 0;
               "Stopped_HMI_Feedback_Tag(1)" := 0;
               "Running_HMI_Feedback_Tag(1)" := 0;
               "Ready_For_Task_HMI_Feedback_Tag(1)" := 0;
               "Cnv_Occupied_HMI_Feedback_Tag(1)" := 0;
               "Shuttle_in_place_HMI_Feedback_Tag(1)" := 0;
               "Current_Task_Type_HMI_Feedback_Tag(1)" := 0;
               "Current_Task_ID_HMI_Feedback_Tag(1)" := 0;
               "SM_State_HMI_Feedback_Tag(1)" := 0;
               "Motor_Speed_Requested_HMI_Feedback_Tag(1)" := 0;
               "Motor_Speed_Actual_HMI_Feedback_Tag(1)" := 0;
           ELSE
               "Same_Cnv" := FALSE;
           END_IF;
           "R_TRIG_DB_2"(CLK := "Same_Cnv");

           IF "R_TRIG_DB_2".Q THEN
               "CNV_ID_HMI_Tag" := 0;
               "CNV_ID_HMI_Tag(1)" := 0;
           END_IF;

           //CHARGE DATA CHANGING CONVEYORS ID
           IF "CNV_ID_HMI_Tag" <> "CNV_ID_HMI_Tag_Old" THEN
               "Screen_DB".Charge_Cnv_Commands := TRUE;
               "CNV_ID_HMI_Tag_Old" := "CNV_ID_HMI_Tag";
           END_IF;

           "R_TRIG_DB_1"(CLK := "Screen_DB".Charge_Cnv_Commands);

           IF "R_TRIG_DB_1".Q THEN
               IF "CNV_ID_HMI_Tag" >= 120001 AND "CNV_ID_HMI_Tag" <= 120301 THEN //ECONVEYOR
                   "Enable_HMI_Tag" := "Control_DB".ECnv_Control.Instruction.Enable;
                   "Mode_Change_HMI_Tag" := "Control_DB".ECnv_Control.Instruction.Mode_Change;
                   "Task_ID_HMI_Tag" := "Control_DB".ECnv_Control.Instruction.Task_ID;
                   "Transfer_To_ID_HMI_Tag" := "Control_DB".ECnv_Control.Instruction.Transfer_To_ID;
                   "Transfer_From_ID_HMI_Tag" := "Control_DB".ECnv_Control.Instruction.Transfer_From_ID;
               ELSIF "CNV_ID_HMI_Tag" >= 100101 AND "CNV_ID_HMI_Tag" <= 100301 THEN //BUFFER CONVEYORS
                   FOR #i := 1 TO 3 DO
                       IF "CNV_ID_HMI_Tag" = "Settings_DB".LCnv_Settings[#i].ID THEN
                           "Enable_HMI_Tag" := "Control_DB".LCnv_Control[#i].Instruction.Enable;
                           "Mode_Change_HMI_Tag" := "Control_DB".LCnv_Control[#i].Instruction.Mode_Change;
                           "Task_ID_HMI_Tag" := "Control_DB".LCnv_Control[#i].Instruction.Task_ID;
                           "Transfer_To_ID_HMI_Tag" := "Control_DB".LCnv_Control[#i].Instruction.Transfer_To_ID;
                           "Transfer_From_ID_HMI_Tag" := "Control_DB".LCnv_Control[#i].Instruction.Transfer_From_ID;
                       END_IF;
                   END_FOR;
               ELSIF "CNV_ID_HMI_Tag" = "Settings_DB".Inbound_Cnv_Settings.ID THEN //INBOUND CONVEYOR
                   "Enable_HMI_Tag" := "Control_DB".Inbound_Cnv.Instruction.Enable;
                   "Mode_Change_HMI_Tag" := "Control_DB".Inbound_Cnv.Instruction.Mode_Change;
                   "Task_ID_HMI_Tag" := "Control_DB".Inbound_Cnv.Instruction.Task_ID;
                   "Transfer_To_ID_HMI_Tag" := "Control_DB".Inbound_Cnv.Instruction.Transfer_To_ID;
                   "Transfer_From_ID_HMI_Tag" := "Control_DB".Inbound_Cnv.Instruction.Transfer_From_ID;
               ELSIF "CNV_ID_HMI_Tag" = "Settings_DB".Outbound_Cnv_Settings.ID THEN //OUTBOUND CONVEYOR
                   "Enable_HMI_Tag" := "Control_DB".Outbound_Cnv.Instruction.Enable;
                   "Mode_Change_HMI_Tag" := "Control_DB".Outbound_Cnv.Instruction.Mode_Change;
                   "Task_ID_HMI_Tag" := "Control_DB".Outbound_Cnv.Instruction.Task_ID;
                   "Transfer_To_ID_HMI_Tag" := "Control_DB".Outbound_Cnv.Instruction.Transfer_To_ID;
                   "Transfer_From_ID_HMI_Tag" := "Control_DB".Outbound_Cnv.Instruction.Transfer_From_ID;
               ELSIF "CNV_ID_HMI_Tag" >= 150101 AND "CNV_ID_HMI_Tag" <= 180101 THEN //POPUP CONVEYORS
                   FOR #i := 1 TO 4 DO
                       "Enable_HMI_Tag" := "Control_DB".PopUp_Cnv[#i].Instruction.Enable;
                       "Mode_Change_HMI_Tag" := "Control_DB".PopUp_Cnv[#i].Instruction.Mode_Change;
                       "Task_ID_HMI_Tag" := "Control_DB".PopUp_Cnv[#i].Instruction.Task_ID;
                       "Transfer_To_ID_HMI_Tag" := "Control_DB".PopUp_Cnv[#i].Instruction.Transfer_To_ID;
                       "Transfer_From_ID_HMI_Tag" := "Control_DB".PopUp_Cnv[#i].Instruction.Transfer_From_ID;
                   END_FOR;
               END_IF;
               "Screen_DB".Charge_Cnv_Commands := 0;
           END_IF;
       END_REGION

       REGION CHARGE DATA FROM HMI (AFTER CHARGE DATA)
           IF NOT "Screen_DB".Charge_Cnv_Commands THEN
               REGION VTD CONVEYOR
                   IF "CNV_ID_HMI_Tag" >= 120001 AND "CNV_ID_HMI_Tag" <= 120301 THEN
                       "EConveyor_Visibility" := TRUE;

                       //Sensors
                       "HMI_CNV_Pallet Detect 1" := "Control_DB".ECnv_Control.Inputs."Pallet Detect 1";
                       "HMI_CNV_Pallet Detect 2" := "Control_DB".ECnv_Control.Inputs."Pallet Detect 2";
                       "HMI_CNV_Sdetect1" := "Control_DB".ECnv_Control.Inputs.Sdetect1;
                       "HMI_CNV_Sdetect2" := "Control_DB".ECnv_Control.Inputs.Sdetect2;

                       //Feedback
                       "Mode_HMI_Feedback_Tag" := "Control_DB".ECnv_Control.Mode;
                       "Enabled_HMI_Feedback_Tag" := "Control_DB".ECnv_Control.Enabled;
                       "Error_HMI_Feedback_Tag" := "Control_DB".ECnv_Control.Error;
                       "Warning_HMI_Feedback_Tag" := "Control_DB".ECnv_Control.Warning;
                       "Stopped_HMI_Feedback_Tag" := "Control_DB".ECnv_Control.Stopped;
                       "Running_HMI_Feedback_Tag" := "Control_DB".ECnv_Control.Running;
                       "Ready_For_Task_HMI_Feedback_Tag" := "Control_DB".ECnv_Control.Ready_For_Task;
                       "Cnv_Occupied_HMI_Feedback_Tag" := "Control_DB".ECnv_Control.Cnv_Occupied;
                       "Shuttle_in_place_HMI_Feedback_Tag" := "Control_DB".ECnv_Control.Shuttle_In_Place;
                       "Current_Task_Type_HMI_Feedback_Tag" := "Control_DB".ECnv_Control.Current_Task_Type;
                       "Current_Task_ID_HMI_Feedback_Tag" := "Control_DB".ECnv_Control.Current_Task_ID;
                       "SM_State_HMI_Feedback_Tag" := "Control_DB".ECnv_Control.SM_State;
                       IF "Control_DB".ECnv_Control.Motor.Forward THEN
                           "Motor_Direction_HMI_Feedback_Tag" := 1;
                       ELSIF "Control_DB".ECnv_Control.Motor.Reverse THEN
                           "Motor_Direction_HMI_Feedback_Tag" := 2;
                       ELSE
                           "Motor_Direction_HMI_Feedback_Tag" := 0;
                       END_IF;
                       "Motor_Speed_Requested_HMI_Feedback_Tag" := "Control_DB".ECnv_Control.Motor.Speed;
                       "Motor_Speed_Actual_HMI_Feedback_Tag" := "Control_DB".ECnv_Control.Motor.Speed_Actual;
                       "Transfer_To_ID_HMI_Tag" := "Control_DB".ECnv_Control.Instruction.Transfer_To_ID;
                       "Transfer_From_ID_HMI_Tag" := "Control_DB".ECnv_Control.Instruction.Transfer_From_ID;

                       //Instructions
                       IF "HMI_DB".ScreenNo = 2 THEN
                           "Control_DB".ECnv_Control.Instruction.Stop := "Stop_HMI_Tag";
                           "Control_DB".ECnv_Control.Instruction.Execute := "Manual_Fwd_HMI_Tag" OR "Manual_Bwd_HMI_Tag";
                           "Control_DB".ECnv_Control.Instruction.Mode_Change := "Mode_Change_HMI_Tag";
                           "Control_DB".ECnv_Control.Instruction.Enable := "Enable_HMI_Tag";
                           IF "Control_DB".ECnv_Control.Mode <> 3 THEN
                               "Control_DB".ECnv_Control.Instruction.Foward := "Manual_Fwd_HMI_Tag";
                               "Control_DB".ECnv_Control.Instruction.Backward := "Manual_Bwd_HMI_Tag";
                               "Control_DB".ECnv_Control.Instruction.Start_Transfer := "Start_Transfer_HMI_Tag";
                               IF "Control_DB".ECnv_Control.Mode = 1 THEN
                                   "Control_DB".ECnv_Control.Instruction.Start_Transfer_Backward := "Transfer_Backward";
                               END_IF;
                               "Control_DB".ECnv_Control.Instruction.Task_ID := "Task_ID_HMI_Tag";
                               IF "CNV_In_Out" THEN // 0 = Inbound, 1 = Outbound
                                   "Control_DB".ECnv_Control.Instruction.Transfer_To_ID := "CNV_ID_HMI_Tag(1)";
                                   "Control_DB".ECnv_Control.Instruction.Transfer_From_ID := 0;
                               ELSE
                                   "Control_DB".ECnv_Control.Instruction.Transfer_To_ID := 0;
                                   "Control_DB".ECnv_Control.Instruction.Transfer_From_ID := "CNV_ID_HMI_Tag(1)";
                               END_IF;
                           END_IF;
                       END_IF;
                   END_IF;
               END_REGION

               REGION BUFFER CONVEYORS
                   FOR #i := 1 TO 3 DO
                       IF "CNV_ID_HMI_Tag" = "Settings_DB".LCnv_Settings[#i].ID THEN
                           //Sensors
                           "HMI_CNV_Pallet Detect 1" := "Control_DB".LCnv_Control[#i].Inputs."Pallet Detect 1";
                           "HMI_CNV_Pallet Detect 2" := "Control_DB".LCnv_Control[#i].Inputs."Pallet Detect 2";
                           "HMI_CNV_Pallet Detect 3" := "Control_DB".LCnv_Control[#i].Inputs."Pallet Detect 3";
                           "HMI_CNV_Sdetect1" := "Control_DB".LCnv_Control[#i].Inputs.Sdetect1;
                           "HMI_CNV_Sdetect2" := "Control_DB".LCnv_Control[#i].Inputs.Sdetect2;
                           "HMI_CNV_SftyPinUp" := "Control_DB".LCnv_Control[#i].Inputs.SftyPinUp;
                           "HMI_CNV_SftyPinDown" := "Control_DB".LCnv_Control[#i].Inputs.SftyPinDown;
                           IF "Control_DB".LCnv_Control[#i].Inputs.SftyPinUp AND NOT "Control_DB".LCnv_Control[#i].Inputs.SftyPinDown THEN
                               "UP_DOWN" := 1;
                           ELSIF NOT "Control_DB".LCnv_Control[#i].Inputs.SftyPinUp AND "Control_DB".LCnv_Control[#i].Inputs.SftyPinDown THEN
                               "UP_DOWN" := 2;
                           ELSE
                               "UP_DOWN" := 0;
                           END_IF;

                           //Feedback
                           "Mode_HMI_Feedback_Tag" := "Control_DB".LCnv_Control[#i].Mode;
                           "Enabled_HMI_Feedback_Tag" := "Control_DB".LCnv_Control[#i].Enabled;
                           "Error_HMI_Feedback_Tag" := "Control_DB".LCnv_Control[#i].Error;
                           "Warning_HMI_Feedback_Tag" := "Control_DB".LCnv_Control[#i].Warning;
                           "Stopped_HMI_Feedback_Tag" := "Control_DB".LCnv_Control[#i].Stopped;
                           "Running_HMI_Feedback_Tag" := "Control_DB".LCnv_Control[#i].Running;
                           "Ready_For_Task_HMI_Feedback_Tag" := "Control_DB".LCnv_Control[#i].Ready_For_Task;
                           "Cnv_Occupied_HMI_Feedback_Tag" := "Control_DB".LCnv_Control[#i].Cnv_Occupied;
                           "Shuttle_in_place_HMI_Feedback_Tag" := "Control_DB".LCnv_Control[#i].Shuttle_In_Place;
                           "Current_Task_Type_HMI_Feedback_Tag" := "Control_DB".LCnv_Control[#i].Current_Task_Type;
                           "Current_Task_ID_HMI_Feedback_Tag" := "Control_DB".LCnv_Control[#i].Current_Task_ID;
                           "SM_State_HMI_Feedback_Tag" := "Control_DB".LCnv_Control[#i].SM_State;
                           IF "Control_DB".LCnv_Control[#i].Motor.Forward THEN
                               "Motor_Direction_HMI_Feedback_Tag" := 1;
                           ELSIF "Control_DB".LCnv_Control[#i].Motor.Reverse THEN
                               "Motor_Direction_HMI_Feedback_Tag" := 2;
                           ELSE
                               "Motor_Direction_HMI_Feedback_Tag" := 0;
                           END_IF;
                           "Motor_Speed_Requested_HMI_Feedback_Tag" := "Control_DB".LCnv_Control[#i].Motor.Speed;
                           "Motor_Speed_Actual_HMI_Feedback_Tag" := "Control_DB".LCnv_Control[#i].Motor.Speed_Actual;
                           "Transfer_To_ID_HMI_Tag" := "Control_DB".LCnv_Control[#i].Instruction.Transfer_To_ID;
                           "Transfer_From_ID_HMI_Tag" := "Control_DB".LCnv_Control[#i].Instruction.Transfer_From_ID;

                           //Instructions
                           IF "HMI_DB".ScreenNo = 2 THEN
                               "Control_DB".LCnv_Control[#i].Instruction.Stop := "Stop_HMI_Tag";
                               "Control_DB".LCnv_Control[#i].Instruction.Execute := "Manual_Fwd_HMI_Tag" OR "Manual_Bwd_HMI_Tag";
                               "Control_DB".LCnv_Control[#i].Instruction.Mode_Change := "Mode_Change_HMI_Tag";
                               "Control_DB".LCnv_Control[#i].Instruction.Enable := "Enable_HMI_Tag";
                               IF "Control_DB".LCnv_Control[#i].Mode <> 3 THEN
                                   "Control_DB".LCnv_Control[#i].Instruction.Foward := "Manual_Fwd_HMI_Tag";
                                   "Control_DB".LCnv_Control[#i].Instruction.Backward := "Manual_Bwd_HMI_Tag";
                                   "Control_DB".LCnv_Control[#i].Instruction.Start_Transfer := "Start_Transfer_HMI_Tag";
                                   IF "Control_DB".LCnv_Control[#i].Mode = 1 THEN
                                       "Control_DB".LCnv_Control[#i].Instruction.Start_Transfer_Backward := "Transfer_Backward";
                                   END_IF;
                                   "Control_DB".LCnv_Control[#i].Safety_Stop_Cnrl.Instruction.Manual_Extend := "Manual_Sfty_Stopper_Up";
                                   "Control_DB".LCnv_Control[#i].Safety_Stop_Cnrl.Instruction.Manual_Retract := "Manual_Sfty_Stopper_Down";
                                   "Control_DB".LCnv_Control[#i].Instruction.Task_ID := "Task_ID_HMI_Tag";
                                   // "Control_DB".LCnv_Control[#i].Instruction.Transfer_To_ID := "Transfer_To_ID_HMI_Tag";
                                   // "Control_DB".LCnv_Control[#i].Instruction.Transfer_From_ID := "Transfer_From_ID_HMI_Tag";
                                   IF "CNV_In_Out" THEN // 0 = Inbound, 1 = Outbound
                                       "Control_DB".LCnv_Control[#i].Instruction.Transfer_To_ID := DINT#120001 + (#i * 100);
                                       "Control_DB".LCnv_Control[#i].Instruction.Transfer_From_ID := 0;
                                   ELSE
                                       "Control_DB".LCnv_Control[#i].Instruction.Transfer_To_ID := 0;
                                       "Control_DB".LCnv_Control[#i].Instruction.Transfer_From_ID := DINT#120001 + (#i * 100);
                                   END_IF;
                               END_IF;
                           END_IF;
                       END_IF;
                   END_FOR;
               END_REGION

               REGION INBOUND CONVEYOR
                   IF "CNV_ID_HMI_Tag" = "Settings_DB".Inbound_Cnv_Settings.ID THEN
                       //Sensors
                       "HMI_CNV_Pallet Detect 1" := "Control_DB".Inbound_Cnv."Inputs"."Pallet Detect 1";
                       "HMI_CNV_Pallet Detect 2" := "Control_DB".Inbound_Cnv.Inputs."Pallet Detect 2";

                       //Feedback
                       "Mode_HMI_Feedback_Tag" := "Control_DB".Inbound_Cnv.Mode;
                       "Enabled_HMI_Feedback_Tag" := "Control_DB".Inbound_Cnv.Enabled;
                       "Error_HMI_Feedback_Tag" := "Control_DB".Inbound_Cnv.Error;
                       "Warning_HMI_Feedback_Tag" := "Control_DB".Inbound_Cnv.Warning;
                       "Stopped_HMI_Feedback_Tag" := "Control_DB".Inbound_Cnv.Stopped;
                       "Running_HMI_Feedback_Tag" := "Control_DB".Inbound_Cnv.Running;
                       "Ready_For_Task_HMI_Feedback_Tag" := "Control_DB".Inbound_Cnv.Ready_For_Task;
                       "Cnv_Occupied_HMI_Feedback_Tag" := "Control_DB".Inbound_Cnv.Cnv_Occupied;
                       "Current_Task_Type_HMI_Feedback_Tag" := "Control_DB".Inbound_Cnv.Current_Task_Type;
                       "Current_Task_ID_HMI_Feedback_Tag" := "Control_DB".Inbound_Cnv.Current_Task_ID;
                       "SM_State_HMI_Feedback_Tag" := "Control_DB".Inbound_Cnv.SM_State;
                       IF "Control_DB".Inbound_Cnv.Motor.Forward THEN
                           "Motor_Direction_HMI_Feedback_Tag" := 1;
                       ELSIF "Control_DB".Inbound_Cnv.Motor.Reverse THEN
                           "Motor_Direction_HMI_Feedback_Tag" := 2;
                       ELSE
                           "Motor_Direction_HMI_Feedback_Tag" := 0;
                       END_IF;
                       "Motor_Speed_Requested_HMI_Feedback_Tag" := "Control_DB".Inbound_Cnv.Motor.Speed;
                       "Motor_Speed_Actual_HMI_Feedback_Tag" := "Control_DB".Inbound_Cnv.Motor.Speed_Actual;
                       "Transfer_To_ID_HMI_Tag" := "Control_DB".Inbound_Cnv.Instruction.Transfer_To_ID;
                       "Transfer_From_ID_HMI_Tag" := "Control_DB".Inbound_Cnv.Instruction.Transfer_From_ID;

                       //Instructions
                       IF "HMI_DB".ScreenNo = 2 THEN
                           "Control_DB".Inbound_Cnv.Instruction.Stop := "Stop_HMI_Tag";
                           "Control_DB".Inbound_Cnv.Instruction.Execute := "Manual_Fwd_HMI_Tag" OR "Manual_Bwd_HMI_Tag";
                           "Control_DB".Inbound_Cnv.Instruction.Mode_Change := "Mode_Change_HMI_Tag";
                           "Control_DB".Inbound_Cnv.Instruction.Enable := "Enable_HMI_Tag";
                           IF "Control_DB".Inbound_Cnv.Mode <> 3 THEN
                               "Control_DB".Inbound_Cnv.Instruction.Foward := "Manual_Fwd_HMI_Tag";
                               "Control_DB".Inbound_Cnv.Instruction.Backward := "Manual_Bwd_HMI_Tag";
                               "Control_DB".Inbound_Cnv.Instruction.Start_Transfer := "Start_Transfer_HMI_Tag";
                               IF "Control_DB".Inbound_Cnv.Mode = 1  THEN
                                   "Control_DB".Inbound_Cnv.Instruction.Start_Transfer_Backward := "Transfer_Backward";
                               END_IF;
                               "Control_DB".Inbound_Cnv.Instruction.Task_ID := "Task_ID_HMI_Tag";
                               "Control_DB".Inbound_Cnv.Instruction.Transfer_To_ID := "Settings_DB".PopUp_Cnv_Settings[1].ID;
                           END_IF;
                       END_IF;
                   END_IF;
               END_REGION

               REGION OUTBOUND CONVEYOR
                   IF "CNV_ID_HMI_Tag" = "Settings_DB".Outbound_Cnv_Settings.ID THEN
                       //Sensors
                       "HMI_CNV_Pallet Detect 1" := "Control_DB".Outbound_Cnv.Inputs."Pallet Detect";

                       //Feedback
                       "Mode_HMI_Feedback_Tag" := "Control_DB".Outbound_Cnv.Mode;
                       "Enabled_HMI_Feedback_Tag" := "Control_DB".Outbound_Cnv.Enabled;
                       "Error_HMI_Feedback_Tag" := "Control_DB".Outbound_Cnv.Error;
                       "Warning_HMI_Feedback_Tag" := "Control_DB".Outbound_Cnv.Warning;
                       "Stopped_HMI_Feedback_Tag" := "Control_DB".Outbound_Cnv.Stopped;
                       "Running_HMI_Feedback_Tag" := "Control_DB".Outbound_Cnv.Running;
                       "Ready_For_Task_HMI_Feedback_Tag" := "Control_DB".Outbound_Cnv.Ready_For_Task;
                       "Cnv_Occupied_HMI_Feedback_Tag" := "Control_DB".Outbound_Cnv.Cnv_Occupied;
                       "Shuttle_in_place_HMI_Feedback_Tag" := "Control_DB".Outbound_Cnv.Shuttle_In_Place;
                       "Current_Task_Type_HMI_Feedback_Tag" := "Control_DB".Outbound_Cnv.Current_Task_Type;
                       "Current_Task_ID_HMI_Feedback_Tag" := "Control_DB".Outbound_Cnv.Current_Task_ID;
                       "SM_State_HMI_Feedback_Tag" := "Control_DB".Outbound_Cnv.SM_State;
                       IF "Control_DB".Outbound_Cnv.Motor.Forward THEN
                           "Motor_Direction_HMI_Feedback_Tag" := 1;
                       ELSIF "Control_DB".Outbound_Cnv.Motor.Reverse THEN
                           "Motor_Direction_HMI_Feedback_Tag" := 2;
                       ELSE
                           "Motor_Direction_HMI_Feedback_Tag" := 0;
                       END_IF;
                       "Motor_Speed_Requested_HMI_Feedback_Tag" := "Control_DB".Outbound_Cnv.Motor.Speed;
                       "Motor_Speed_Actual_HMI_Feedback_Tag" := "Control_DB".Outbound_Cnv.Motor.Speed_Actual;
                       "Transfer_To_ID_HMI_Tag" := "Control_DB".Outbound_Cnv.Instruction.Transfer_To_ID;
                       "Transfer_From_ID_HMI_Tag" := "Control_DB".Outbound_Cnv.Instruction.Transfer_From_ID;

                       //Instructions
                       IF "HMI_DB".ScreenNo = 2 THEN
                           "Control_DB".Outbound_Cnv.Instruction.Stop := "Stop_HMI_Tag";
                           "Control_DB".Outbound_Cnv.Instruction.Execute := "Manual_Fwd_HMI_Tag" OR "Manual_Bwd_HMI_Tag";
                           "Control_DB".Outbound_Cnv.Instruction.Mode_Change := "Mode_Change_HMI_Tag";
                           "Control_DB".Outbound_Cnv.Instruction.Enable := "Enable_HMI_Tag";
                           IF "Control_DB".Outbound_Cnv.Mode <> 3 THEN
                               "Control_DB".Outbound_Cnv.Instruction.Foward := "Manual_Fwd_HMI_Tag";
                               "Control_DB".Outbound_Cnv.Instruction.Backward := "Manual_Bwd_HMI_Tag";
                               "Control_DB".Outbound_Cnv.Instruction.Start_Transfer := "Start_Transfer_HMI_Tag";
                               IF "Control_DB".Outbound_Cnv.Mode = 1 THEN
                                   "Control_DB".Outbound_Cnv.Instruction.Start_Transfer_Backward := "Transfer_Backward";
                               END_IF;
                               "Control_DB".Outbound_Cnv.Instruction.Task_ID := "Task_ID_HMI_Tag";
                               "Control_DB".Outbound_Cnv.Instruction.Transfer_From_ID := "Settings_DB".PopUp_Cnv_Settings[4].ID;
                           END_IF;
                       END_IF;
                   END_IF;
               END_REGION

               REGION POPUP CONVEYORS
                   IF "CNV_ID_HMI_Tag" = "Settings_DB".PopUp_Cnv_Settings[1].ID THEN
                       "HMI_CNV_Pallet Detect 1" := "PopUp Conveyor 1 - Pallet sensor";
                       "HMI_CNV_Pallet Detect 2" := "Pick Station";
                   ELSIF "CNV_ID_HMI_Tag" = "Settings_DB".PopUp_Cnv_Settings[2].ID THEN
                       "HMI_CNV_Pallet Detect 1" := "PopUp Conveyor 2 - Pallet Present 1";
                       "HMI_CNV_Pallet Detect 2" := "PopUp Conveyor 2 - Pallet present 2";
                       "HMI_CNV_Pallet Detect 3" := "PopUp Conveyor 2 - Pallet present 3";
                       "HMI_CNV_Pallet Detect 4" := "PopUp Conveyor 2 - Pallet present 4";
                       "HMI_CNV_Pallet Detect 5" := "PopUp Conveyor 2 - Pallet present 5";
                   ELSIF "CNV_ID_HMI_Tag" = "Settings_DB".PopUp_Cnv_Settings[3].ID THEN
                       "HMI_CNV_Pallet Detect 1" := "PopUp Conveyor 3 - Pallet present 1";
                   ELSIF "CNV_ID_HMI_Tag" = "Settings_DB".PopUp_Cnv_Settings[4].ID THEN
                       "HMI_CNV_Pallet Detect 1" := "PopUp Conveyor 4 - Pallet present 1";
                       "HMI_CNV_Pallet Detect 2" := "Pick Station";
                   END_IF;
                   FOR #i := 1 TO 4 DO
                       IF "CNV_ID_HMI_Tag" = "Settings_DB".PopUp_Cnv_Settings[#i].ID THEN
                           //Sensors
                           IF "Control_DB".PopUp_Cnv[#i].Inputs."Lift Up" AND NOT "Control_DB".PopUp_Cnv[#i].Inputs."Lift Down" THEN
                               "UP_DOWN" := 1;
                           ELSIF NOT "Control_DB".PopUp_Cnv[#i].Inputs."Lift Up" AND "Control_DB".PopUp_Cnv[#i].Inputs."Lift Down" THEN
                               "UP_DOWN" := 2;
                           ELSE
                               "UP_DOWN" := 0;
                           END_IF;
                           IF "CNV_ID_HMI_Tag" = "Settings_DB".PopUp_Cnv_Settings[#i].ID THEN
                               //Feedback
                               "Mode_HMI_Feedback_Tag" := "Control_DB".PopUp_Cnv[#i].Mode;
                               "Enabled_HMI_Feedback_Tag" := "Control_DB".PopUp_Cnv[#i].Enabled;
                               "Error_HMI_Feedback_Tag" := "Control_DB".PopUp_Cnv[#i].Error;
                               "Warning_HMI_Feedback_Tag" := "Control_DB".PopUp_Cnv[#i].Warning;
                               "Stopped_HMI_Feedback_Tag" := "Control_DB".PopUp_Cnv[#i].Stopped;
                               "Running_HMI_Feedback_Tag" := "Control_DB".PopUp_Cnv[#i].Running;
                               "Ready_For_Task_HMI_Feedback_Tag" := "Control_DB".PopUp_Cnv[#i].Ready_For_Task;
                               "Cnv_Occupied_HMI_Feedback_Tag" := "Control_DB".PopUp_Cnv[#i].Cnv_Occupied;
                               "Current_Task_Type_HMI_Feedback_Tag" := "Control_DB".PopUp_Cnv[#i].Current_Task_Type;
                               "Current_Task_ID_HMI_Feedback_Tag" := "Control_DB".PopUp_Cnv[#i].Current_Task_ID;
                               "SM_State_HMI_Feedback_Tag" := "Control_DB".PopUp_Cnv[#i].SM_State;
                               "Transfer_To_ID_HMI_Tag" := "Control_DB".PopUp_Cnv[#i].Instruction.Transfer_To_ID;
                               "Transfer_From_ID_HMI_Tag" := "Control_DB".PopUp_Cnv[#i].Instruction.Transfer_From_ID;
                               IF "Control_DB".PopUp_Cnv[#i].Roller_Motor.Status.%X0 THEN
                                   IF "Control_DB".PopUp_Cnv[#i].Roller_Motor.Forward THEN
                                       "Motor_Direction_HMI_Feedback_Tag" := 1;
                                   ELSIF "Control_DB".PopUp_Cnv[#i].Roller_Motor.Reverse THEN
                                       "Motor_Direction_HMI_Feedback_Tag" := 2;
                                   ELSE
                                       "Motor_Direction_HMI_Feedback_Tag" := 0;
                                   END_IF;
                                   "Motor_Speed_Requested_HMI_Feedback_Tag" := REAL_TO_UINT("Control_DB".PopUp_Cnv[#i].Roller_Motor.Speed);
                                   "Motor_Speed_Actual_HMI_Feedback_Tag" := REAL_TO_UINT("Control_DB".PopUp_Cnv[#i].Roller_Motor.Speed_Actual);
                               ELSIF "Control_DB".PopUp_Cnv[#i].Chain_Motor.Status.%X0 = 1 THEN
                                   IF "Control_DB".PopUp_Cnv[#i].Chain_Motor.Forward THEN
                                       "Motor_Direction_HMI_Feedback_Tag" := 1;
                                   ELSIF "Control_DB".PopUp_Cnv[#i].Chain_Motor.Reverse THEN
                                       "Motor_Direction_HMI_Feedback_Tag" := 2;
                                   ELSE
                                       "Motor_Direction_HMI_Feedback_Tag" := 0;
                                   END_IF;
                                   "Motor_Speed_Requested_HMI_Feedback_Tag" := REAL_TO_UINT("Control_DB".PopUp_Cnv[#i].Chain_Motor.Speed);
                                   "Motor_Speed_Actual_HMI_Feedback_Tag" := REAL_TO_UINT("Control_DB".PopUp_Cnv[#i].Chain_Motor.Speed_Actual);
                               ELSIF "Control_DB".PopUp_Cnv[#i].Lift_Motor.Status.%X0 = 1 THEN
                                   IF "Control_DB".PopUp_Cnv[#i].Lift_Motor.Forward THEN
                                       "Motor_Direction_HMI_Feedback_Tag" := 1;
                                   ELSIF "Control_DB".PopUp_Cnv[#i].Lift_Motor.Reverse THEN
                                       "Motor_Direction_HMI_Feedback_Tag" := 2;
                                   ELSE
                                       "Motor_Direction_HMI_Feedback_Tag" := 0;
                                   END_IF;
                                   "Motor_Speed_Requested_HMI_Feedback_Tag" := REAL_TO_UINT("Control_DB".PopUp_Cnv[#i].Lift_Motor.Speed);
                                   "Motor_Speed_Actual_HMI_Feedback_Tag" := REAL_TO_UINT("Control_DB".PopUp_Cnv[#i].Lift_Motor.Speed_Actual);
                               END_IF;

                               //Instructions
                               IF "HMI_DB".ScreenNo = 2 THEN
                                   "Control_DB".PopUp_Cnv[#i].Instruction.Stop := "Stop_HMI_Tag";
                                   "Control_DB".PopUp_Cnv[#i].Instruction.Execute := "Manual_Fwd_HMI_Tag" OR "Manual_Bwd_HMI_Tag";
                                   "Control_DB".PopUp_Cnv[#i].Instruction.Mode_Change := "Mode_Change_HMI_Tag";
                                   "Control_DB".PopUp_Cnv[#i].Instruction.Enable := "Enable_HMI_Tag";
                                   IF "Control_DB".PopUp_Cnv[#i].Mode <> 3 THEN
                                       IF "Control_DB".PopUp_Cnv[#i].Inputs."Lift Up" THEN
                                           "Control_DB".PopUp_Cnv[#i].Instruction.Roller_Fwd := "Manual_Fwd_HMI_Tag";
                                           "Control_DB".PopUp_Cnv[#i].Instruction.Roller_Bwd := "Manual_Bwd_HMI_Tag";
                                       ELSIF "Control_DB".PopUp_Cnv[#i].Inputs."Lift Down" THEN
                                           "Control_DB".PopUp_Cnv[#i].Instruction.Chain_Fwd := "Manual_Fwd_HMI_Tag";
                                           "Control_DB".PopUp_Cnv[#i].Instruction.Chain_Bwd := "Manual_Bwd_HMI_Tag";
                                       END_IF;
                                       "Control_DB".PopUp_Cnv[#i].Instruction.Start_Transfer := "Start_Transfer_HMI_Tag";
                                       IF "Control_DB".PopUp_Cnv[#i].Mode = 1 THEN
                                           "Control_DB".PopUp_Cnv[#i].Instruction.Start_Transfer_Backward := "Transfer_Backward";
                                       END_IF;
                                       "Control_DB".PopUp_Cnv[#i].Instruction.Lift_Up := "Manual_Sfty_Stopper_Up";
                                       "Control_DB".PopUp_Cnv[#i].Instruction.Lift_Down := "Manual_Sfty_Stopper_Down";
                                       "Control_DB".PopUp_Cnv[#i].Instruction.Task_ID := "Task_ID_HMI_Tag";
                                       CASE #i OF
                                           1:
                                               IF "CNV_In_Out" AND "Control_DB".PopUp_Cnv[1].Inputs."Lift Up" THEN // 0 = Inbound, 1 = Outbound
                                                   "Control_DB".PopUp_Cnv[#i].Instruction.Transfer_To_ID := "Settings_DB".PopUp_Cnv_Settings[2].ID;
                                                   "Control_DB".PopUp_Cnv[#i].Instruction.Transfer_From_ID := 0;
                                               ELSIF NOT "CNV_In_Out" AND "Control_DB".PopUp_Cnv[1].Inputs."Lift Down" AND NOT "Pick Station" THEN // 0 = Inbound, 1 = Outbound
                                                   "Control_DB".PopUp_Cnv[#i].Instruction.Transfer_To_ID := 0;
                                                   "Control_DB".PopUp_Cnv[#i].Instruction.Transfer_From_ID := "Settings_DB".Pick_Cnv_Settings.ID;
                                               ELSIF NOT "CNV_In_Out" AND "Control_DB".PopUp_Cnv[1].Inputs."Lift Up" THEN // 0 = Inbound, 1 = Outbound
                                                   "Control_DB".PopUp_Cnv[#i].Instruction.Transfer_To_ID := 0;
                                                   "Control_DB".PopUp_Cnv[#i].Instruction.Transfer_From_ID := "Settings_DB".Inbound_Cnv_Settings.ID;
                                               ELSE
                                                   "Control_DB".PopUp_Cnv[#i].Instruction.Transfer_To_ID := 0;
                                                   "Control_DB".PopUp_Cnv[#i].Instruction.Transfer_From_ID := 0;
                                               END_IF;

                                           2:
                                               IF NOT "CNV_In_Out" AND "Control_DB".PopUp_Cnv[2].Inputs."Lift Up" THEN // UP
                                                   "Control_DB".PopUp_Cnv[#i].Instruction.Transfer_To_ID := 0;
                                                   "Control_DB".PopUp_Cnv[#i].Instruction.Transfer_From_ID := "Settings_DB".PopUp_Cnv_Settings[1].ID;
                                               ELSIF NOT "CNV_In_Out" AND "Control_DB".PopUp_Cnv[2].Inputs."Lift Down" THEN //DOWN
                                                   "Control_DB".PopUp_Cnv[#i].Instruction.Transfer_To_ID := 0;
                                                   "Control_DB".PopUp_Cnv[#i].Instruction.Transfer_From_ID := "Settings_DB".ECnv_Settings.ID;
                                               ELSIF "CNV_In_Out" AND "Control_DB".PopUp_Cnv[2].Inputs."Lift Down" AND NOT "VTD_POPUP2" THEN //DOWN
                                                   "Control_DB".PopUp_Cnv[#i].Instruction.Transfer_To_ID := "Settings_DB".ECnv_Settings.ID;
                                                   "Control_DB".PopUp_Cnv[#i].Instruction.Transfer_From_ID := 0;
                                               ELSIF "CNV_In_Out" AND "Control_DB".PopUp_Cnv[2].Inputs."Lift Down" AND "VTD_POPUP2" THEN //DOWN
                                                   "Control_DB".PopUp_Cnv[#i].Instruction.Transfer_To_ID := "Settings_DB".PopUp_Cnv_Settings[3].ID;
                                                   "Control_DB".PopUp_Cnv[#i].Instruction.Transfer_From_ID := 0;
                                               ELSE
                                                   "Control_DB".PopUp_Cnv[#i].Instruction.Transfer_To_ID := 0;
                                                   "Control_DB".PopUp_Cnv[#i].Instruction.Transfer_From_ID := 0;
                                               END_IF;

                                           3:
                                               IF NOT "CNV_In_Out" AND "Control_DB".PopUp_Cnv[3].Inputs."Lift Down" THEN //inbound chain
                                                   "Control_DB".PopUp_Cnv[#i].Instruction.Transfer_To_ID := 0;
                                                   "Control_DB".PopUp_Cnv[#i].Instruction.Transfer_From_ID := "Settings_DB".PopUp_Cnv_Settings[2].ID;
                                               ELSIF "CNV_In_Out" AND "Control_DB".PopUp_Cnv[3].Inputs."Lift Up" THEN 
                                                   "Control_DB".PopUp_Cnv[#i].Instruction.Transfer_To_ID := "Settings_DB".PopUp_Cnv_Settings[4].ID;
                                                   "Control_DB".PopUp_Cnv[#i].Instruction.Transfer_From_ID := 0;
                                               ELSE
                                                   "Control_DB".PopUp_Cnv[#i].Instruction.Transfer_To_ID := 0;
                                                   "Control_DB".PopUp_Cnv[#i].Instruction.Transfer_From_ID := 0;
                                               END_IF;

                                           4:
                                               IF "CNV_In_Out" AND "Control_DB".PopUp_Cnv[4].Inputs."Lift Up" THEN // 0 = Inbound, 1 = Outbound
                                                   "Control_DB".PopUp_Cnv[#i].Instruction.Transfer_To_ID := "Settings_DB".Outbound_Cnv_Settings.ID;
                                                   "Control_DB".PopUp_Cnv[#i].Instruction.Transfer_From_ID := 0;
                                               ELSIF "CNV_In_Out" AND "Control_DB".PopUp_Cnv[4].Inputs."Lift Down" AND "Pick Station" THEN // 0 = Inbound, 1 = Outbound
                                                   "Control_DB".PopUp_Cnv[#i].Instruction.Transfer_To_ID := "Settings_DB".Pick_Cnv_Settings.ID;
                                                   "Control_DB".PopUp_Cnv[#i].Instruction.Transfer_From_ID := 0;
                                               ELSIF NOT "CNV_In_Out" AND "Control_DB".PopUp_Cnv[4].Inputs."Lift Up" THEN // 0 = Inbound, 1 = Outbound
                                                   "Control_DB".PopUp_Cnv[#i].Instruction.Transfer_To_ID := 0;
                                                   "Control_DB".PopUp_Cnv[#i].Instruction.Transfer_From_ID := "Settings_DB".PopUp_Cnv_Settings[3].ID;
                                               ELSE
                                                   "Control_DB".PopUp_Cnv[#i].Instruction.Transfer_To_ID := 0;
                                                   "Control_DB".PopUp_Cnv[#i].Instruction.Transfer_From_ID := 0;
                                               END_IF;
                                       END_CASE;
                                   END_IF;
                               END_IF;
                           END_IF;
                       END_IF;
                   END_FOR;
               END_REGION

               REGION PICK CONVEYOR
                   IF "CNV_ID_HMI_Tag" = "Settings_DB".Pick_Cnv_Settings.ID THEN
                       //Sensors
                       "HMI_CNV_Pallet Detect 1" := "Control_DB".Pick_Station.Cnv_Occupied;

                       //Feedback
                       "Mode_HMI_Feedback_Tag" := "Control_DB".Pick_Station.Mode;
                       "Enabled_HMI_Feedback_Tag" := "Control_DB".Pick_Station.Enabled;
                       "Error_HMI_Feedback_Tag" := "Control_DB".Pick_Station.Error;
                       "Warning_HMI_Feedback_Tag" := "Control_DB".Pick_Station.Warning;
                       "Stopped_HMI_Feedback_Tag" := "Control_DB".Pick_Station.Stopped;
                       "Running_HMI_Feedback_Tag" := "Control_DB".Pick_Station.Running;
                       "Ready_For_Task_HMI_Feedback_Tag" := "Control_DB".Pick_Station.Ready_For_Task;
                       "Cnv_Occupied_HMI_Feedback_Tag" := "Control_DB".Pick_Station.Cnv_Occupied;
                       // "Shuttle_in_place_HMI_Feedback_Tag" := "Control_DB".Pick_Station.Shuttle_In_Place;
                       "Current_Task_Type_HMI_Feedback_Tag" := "Control_DB".Pick_Station.Current_Task_Type;
                       "Current_Task_ID_HMI_Feedback_Tag" := "Control_DB".Pick_Station.Current_Task_ID;
                       "SM_State_HMI_Feedback_Tag" := "Control_DB".Pick_Station.SM_State;
                       IF "Control_DB".Pick_Station.Motor.Forward THEN
                           "Motor_Direction_HMI_Feedback_Tag" := 1;
                       ELSIF "Control_DB".Pick_Station.Motor.Reverse THEN
                           "Motor_Direction_HMI_Feedback_Tag" := 2;
                       ELSE
                           "Motor_Direction_HMI_Feedback_Tag" := 0;
                       END_IF;
                       "Motor_Speed_Requested_HMI_Feedback_Tag" := "Control_DB".Pick_Station.Motor.Speed;
                       "Motor_Speed_Actual_HMI_Feedback_Tag" := "Control_DB".Pick_Station.Motor.Speed_Actual;
                       "Transfer_To_ID_HMI_Tag" := "Control_DB".Pick_Station.Instruction.Transfer_To_ID;
                       "Transfer_From_ID_HMI_Tag" := "Control_DB".Pick_Station.Instruction.Transfer_From_ID;

                       //Instructions
                       IF "HMI_DB".ScreenNo = 2 THEN
                           "Control_DB".Pick_Station.Instruction.Stop := "Stop_HMI_Tag";
                           "Control_DB".Pick_Station.Instruction.Execute := "Manual_Fwd_HMI_Tag" OR "Manual_Bwd_HMI_Tag";
                           "Control_DB".Pick_Station.Instruction.Mode_Change := "Mode_Change_HMI_Tag";
                           "Control_DB".Pick_Station.Instruction.Enable := "Enable_HMI_Tag";
                           IF "Control_DB".Pick_Station.Mode <> 3 THEN
                               "Control_DB".Pick_Station.Instruction.Foward := "Manual_Fwd_HMI_Tag";
                               "Control_DB".Pick_Station.Instruction.Backward := "Manual_Bwd_HMI_Tag";
                               "Control_DB".Pick_Station.Instruction.Start_Transfer := "Start_Transfer_HMI_Tag";
                               IF "Control_DB".Pick_Station.Mode = 1 THEN
                                   "Control_DB".Pick_Station.Instruction.Start_Transfer_Backward := "Transfer_Backward";
                               END_IF;
                               "Control_DB".Pick_Station.Instruction.Task_ID := "Task_ID_HMI_Tag";
                               "Control_DB".Pick_Station.Instruction.Transfer_From_ID := "Settings_DB".PopUp_Cnv_Settings[4].ID;
                               "Control_DB".Pick_Station.Instruction.Transfer_To_ID := "Settings_DB".PopUp_Cnv_Settings[1].ID;
                           END_IF;
                       END_IF;
                   END_IF;
               END_REGION
           END_IF;
       END_REGION
   END_REGION


   REGION Assign Conveyor 2
       REGION Charge DATA to HMI
           //CHARGE DATA CHANGING CONVEYORS ID
           IF "CNV_ID_HMI_Tag(1)" <> "CNV_ID_HMI_Tag(1)_Old" THEN
               "Screen_DB".Charge_Cnv_Commands := TRUE;
               "CNV_ID_HMI_Tag(1)_Old" := "CNV_ID_HMI_Tag(1)";
           END_IF;

           "R_TRIG_DB_7"(CLK := "Screen_DB".Charge_Cnv_Commands);

           IF "R_TRIG_DB_7".Q THEN
               IF "CNV_ID_HMI_Tag(1)" >= 120001 AND "CNV_ID_HMI_Tag(1)" <= 120301 THEN //ECONVEYOR
                   "Enable_HMI_Tag(1)" := "Control_DB".ECnv_Control.Instruction.Enable;
                   "Mode_Change_HMI_Tag(1)" := "Control_DB".ECnv_Control.Instruction.Mode_Change;
                   "Task_ID_HMI_Tag(1)" := "Control_DB".ECnv_Control.Instruction.Task_ID;
                   "Transfer_To_ID_HMI_Tag(1)" := "Control_DB".ECnv_Control.Instruction.Transfer_To_ID;
                   "Transfer_From_ID_HMI_Tag(1)" := "Control_DB".ECnv_Control.Instruction.Transfer_From_ID;
               ELSIF "CNV_ID_HMI_Tag" >= 100101 AND "CNV_ID_HMI_Tag" <= 100301 THEN //BUFFER CONVEYORS
                   FOR #i := 1 TO 3 DO
                       IF "CNV_ID_HMI_Tag(1)" = "Settings_DB".LCnv_Settings[#i].ID THEN
                           "Enable_HMI_Tag(1)" := "Control_DB".LCnv_Control[#i].Instruction.Enable;
                           "Mode_Change_HMI_Tag(1)" := "Control_DB".LCnv_Control[#i].Instruction.Mode_Change;
                           "Task_ID_HMI_Tag(1)" := "Control_DB".LCnv_Control[#i].Instruction.Task_ID;
                           "Transfer_To_ID_HMI_Tag(1)" := "Control_DB".LCnv_Control[#i].Instruction.Transfer_To_ID;
                           "Transfer_From_ID_HMI_Tag(1)" := "Control_DB".LCnv_Control[#i].Instruction.Transfer_From_ID;
                       END_IF;
                   END_FOR;
               ELSIF "CNV_ID_HMI_Tag(1)" = "Settings_DB".Inbound_Cnv_Settings.ID THEN //INBOUND CONVEYOR
                   "Enable_HMI_Tag(1)" := "Control_DB".Inbound_Cnv.Instruction.Enable;
                   "Mode_Change_HMI_Tag(1)" := "Control_DB".Inbound_Cnv.Instruction.Mode_Change;
                   "Task_ID_HMI_Tag(1)" := "Control_DB".Inbound_Cnv.Instruction.Task_ID;
                   "Transfer_To_ID_HMI_Tag(1)" := "Control_DB".Inbound_Cnv.Instruction.Transfer_To_ID;
                   "Transfer_From_ID_HMI_Tag(1)" := "Control_DB".Inbound_Cnv.Instruction.Transfer_From_ID;
               ELSIF "CNV_ID_HMI_Tag(1)" = "Settings_DB".Outbound_Cnv_Settings.ID THEN //OUTBOUND CONVEYOR
                   "Enable_HMI_Tag(1)" := "Control_DB".Outbound_Cnv.Instruction.Enable;
                   "Mode_Change_HMI_Tag(1)" := "Control_DB".Outbound_Cnv.Instruction.Mode_Change;
                   "Task_ID_HMI_Tag(1)" := "Control_DB".Outbound_Cnv.Instruction.Task_ID;
                   "Transfer_To_ID_HMI_Tag(1)" := "Control_DB".Outbound_Cnv.Instruction.Transfer_To_ID;
                   "Transfer_From_ID_HMI_Tag(1)" := "Control_DB".Outbound_Cnv.Instruction.Transfer_From_ID;
               ELSIF "CNV_ID_HMI_Tag(1)" >= 150101 AND "CNV_ID_HMI_Tag(1)" <= 180101 THEN //POPUP CONVEYORS
                   FOR #i := 1 TO 4 DO
                       "Enable_HMI_Tag(1)" := "Control_DB".PopUp_Cnv[#i].Instruction.Enable;
                       "Mode_Change_HMI_Tag(1)" := "Control_DB".PopUp_Cnv[#i].Instruction.Mode_Change;
                       "Task_ID_HMI_Tag(1)" := "Control_DB".PopUp_Cnv[#i].Instruction.Task_ID;
                       "Transfer_To_ID_HMI_Tag(1)" := "Control_DB".PopUp_Cnv[#i].Instruction.Transfer_To_ID;
                       "Transfer_From_ID_HMI_Tag(1)" := "Control_DB".PopUp_Cnv[#i].Instruction.Transfer_From_ID;
                   END_FOR;
               END_IF;
               "Screen_DB".Charge_Cnv_Commands := 0;
           END_IF;
       END_REGION

       REGION CHARGE DATA FROM HMI (AFTER CHARGE DATA)
           IF NOT "Screen_DB".Charge_Cnv_Commands THEN
               REGION VTD CONVEYOR
                   IF "CNV_ID_HMI_Tag(1)" >= 120001 AND "CNV_ID_HMI_Tag(1)" <= 120301 THEN
                       "BConveyor_Visibility" := TRUE;

                       //Sensors
                       "HMI_CNV_Pallet Detect 1(1)" := "Control_DB".ECnv_Control.Inputs."Pallet Detect 1";
                       "HMI_CNV_Pallet Detect 2(1)" := "Control_DB".ECnv_Control.Inputs."Pallet Detect 2";
                       "HMI_CNV_Sdetect1(1)" := "Control_DB".ECnv_Control.Inputs.Sdetect1;
                       "HMI_CNV_Sdetect2(1)" := "Control_DB".ECnv_Control.Inputs.Sdetect2;

                       //Feedback
                       "Mode_HMI_Feedback_Tag(1)" := "Control_DB".ECnv_Control.Mode;
                       "Enabled_HMI_Feedback_Tag(1)" := "Control_DB".ECnv_Control.Enabled;
                       "Error_HMI_Feedback_Tag(1)" := "Control_DB".ECnv_Control.Error;
                       "Warning_HMI_Feedback_Tag(1)" := "Control_DB".ECnv_Control.Warning;
                       "Stopped_HMI_Feedback_Tag(1)" := "Control_DB".ECnv_Control.Stopped;
                       "Running_HMI_Feedback_Tag(1)" := "Control_DB".ECnv_Control.Running;
                       "Ready_For_Task_HMI_Feedback_Tag(1)" := "Control_DB".ECnv_Control.Ready_For_Task;
                       "Cnv_Occupied_HMI_Feedback_Tag(1)" := "Control_DB".ECnv_Control.Cnv_Occupied;
                       "Shuttle_in_place_HMI_Feedback_Tag(1)" := "Control_DB".ECnv_Control.Shuttle_In_Place;
                       "Current_Task_Type_HMI_Feedback_Tag(1)" := "Control_DB".ECnv_Control.Current_Task_Type;
                       "Current_Task_ID_HMI_Feedback_Tag(1)" := "Control_DB".ECnv_Control.Current_Task_ID;
                       "SM_State_HMI_Feedback_Tag(1)" := "Control_DB".ECnv_Control.SM_State;
                       IF "Control_DB".ECnv_Control.Motor.Forward THEN
                           "Motor_Direction_HMI_Feedback_Tag(1)" := 1;
                       ELSIF "Control_DB".ECnv_Control.Motor.Reverse THEN
                           "Motor_Direction_HMI_Feedback_Tag(1)" := 2;
                       ELSE
                           "Motor_Direction_HMI_Feedback_Tag(1)" := 0;
                       END_IF;
                       "Motor_Speed_Requested_HMI_Feedback_Tag(1)" := "Control_DB".ECnv_Control.Motor.Speed;
                       "Motor_Speed_Actual_HMI_Feedback_Tag(1)" := "Control_DB".ECnv_Control.Motor.Speed_Actual;
                       "Transfer_To_ID_HMI_Tag(1)" := "Control_DB".ECnv_Control.Instruction.Transfer_To_ID;
                       "Transfer_From_ID_HMI_Tag(1)" := "Control_DB".ECnv_Control.Instruction.Transfer_From_ID;

                       //Instructions
                       IF "HMI_DB".ScreenNo = 2 THEN
                           "Control_DB".ECnv_Control.Instruction.Stop := "Stop_HMI_Tag(1)";
                           "Control_DB".ECnv_Control.Instruction.Mode_Change := "Mode_Change_HMI_Tag(1)";
                           "Control_DB".ECnv_Control.Instruction.Enable := "Enable_HMI_Tag(1)";
                           IF "Control_DB".ECnv_Control.Mode <> 3 THEN
                               "Control_DB".ECnv_Control.Instruction.Task_ID := "Task_ID_HMI_Tag(1)";
                               IF "CNV_In_Out(1)" THEN // 0 = Inbound, 1 = Outbound
                                   "Control_DB".ECnv_Control.Instruction.Transfer_To_ID := "CNV_ID_HMI_Tag";
                                   "Control_DB".ECnv_Control.Instruction.Transfer_From_ID := 0;
                               ELSE
                                   "Control_DB".ECnv_Control.Instruction.Transfer_To_ID := 0;
                                   "Control_DB".ECnv_Control.Instruction.Transfer_From_ID := "CNV_ID_HMI_Tag";
                               END_IF;
                               "Control_DB".ECnv_Control.Instruction.Foward := "Manual_Fwd_HMI_Tag(1)";
                               "Control_DB".ECnv_Control.Instruction.Backward := "Manual_Bwd_HMI_Tag(1)";
                               "Control_DB".ECnv_Control.Instruction.Start_Transfer := "Start_Transfer_HMI_Tag(1)";
                               IF "Control_DB".ECnv_Control.Mode = 1 THEN
                                   "Control_DB".ECnv_Control.Instruction.Start_Transfer_Backward := "Transfer_Backward(1)";
                               END_IF;
                           END_IF;
                       END_IF;
                   END_IF;
               END_REGION

               REGION BUFFER CONVEYORS
                   FOR #i := 1 TO 3 DO
                       IF "CNV_ID_HMI_Tag(1)" = "Settings_DB".LCnv_Settings[#i].ID THEN
                           //Sensors
                           "HMI_CNV_Pallet Detect 1(1)" := "Control_DB".LCnv_Control[#i].Inputs."Pallet Detect 1";
                           "HMI_CNV_Pallet Detect 2(1)" := "Control_DB".LCnv_Control[#i].Inputs."Pallet Detect 2";
                           "HMI_CNV_Pallet Detect 3(1)" := "Control_DB".LCnv_Control[#i].Inputs."Pallet Detect 3";
                           "HMI_CNV_Sdetect1(1)" := "Control_DB".LCnv_Control[#i].Inputs.Sdetect1;
                           "HMI_CNV_Sdetect2(1)" := "Control_DB".LCnv_Control[#i].Inputs.Sdetect2;
                           "HMI_CNV_SftyPinUp(1)" := "Control_DB".LCnv_Control[#i].Inputs.SftyPinUp;
                           "HMI_CNV_SftyPinDown(1)" := "Control_DB".LCnv_Control[#i].Inputs.SftyPinDown;
                           IF "Control_DB".LCnv_Control[#i].Inputs.SftyPinUp AND NOT "Control_DB".LCnv_Control[#i].Inputs.SftyPinDown THEN
                               "UP_DOWN(1)" := 1;
                           ELSIF NOT "Control_DB".LCnv_Control[#i].Inputs.SftyPinUp AND "Control_DB".LCnv_Control[#i].Inputs.SftyPinDown THEN
                               "UP_DOWN(1)" := 2;
                           ELSE
                               "UP_DOWN(1)" := 0;
                           END_IF;

